(* IEC 61131-3 sources: JingjiangMoonbox/Application/Application/任务列表/CommTask/PRG_COMM, 7 files *)

(* ---- Action_gLink_II_Input.st ---- *)
(*@CES
Name=Action_gLink_II_Input
Type=Action
TypeGuid=8ac092e5-3128-4e26-9e7e-11016c6684f2
Guid=1dfcb6d0-4c04-4e1c-b741-2802373335cf
HasDeclaration=False
HasImplementation=True
*)
{DECLARATION}

{IMPLEMENTATION}
FOR iN:=1 TO MAX_UNIT_NUM BY 1 DO
	pstStUnitParam_Save:= ADR(g_stStSysParam.astStUnitParam_Save[iN]);
	pstStUnitParam_UnSave:= ADR(g_stStSysParam.astStUnitParam_UnSave[iN]);
	//xi.hy2026.5.9.114008
	pstStRSVUnitParam_UnSave:=ADR(g_stStSysParam.astStRSV_UnitParam_UnSave[iN]);

	astStParam_Mailbox_snd[iN].dwSemaphore:= SEMA_DOWNLOAD;
	astStParam_Mailbox_snd[iN].iGateSa:= pstStUnitParam_Save^.iGateSa;
	astStParam_Mailbox_snd[iN].iGateSaEx:= pstStUnitParam_Save^.iGateSaEx;
	astStParam_Mailbox_snd[iN].rAdjust_V:= pstStUnitParam_Save^.rAdj_V;
	astStParam_Mailbox_snd[iN].rAdjust_H:= pstStUnitParam_Save^.rAdj_H;
	astStParam_Mailbox_snd[iN].dwFlag_Ctl:= pstStUnitParam_Save^.dwFlag_Ctl;
	astStParam_Mailbox_snd[iN].dwFlag_Sts:= pstStUnitParam_Save^.dwFlag_Sts;
	//2026.04.08.193624//wButtonFun_Lamp赋值
	pstStUnitParam_Save^.wButtonFun_Lamp.0:=g_astStIOMap_Axis_FE[iN].o_xLamp_Linkage;
	pstStUnitParam_Save^.wButtonFun_Lamp.3:=g_astStIOMap_Axis_FE[iN].o_xLamp_Inch;
	pstStUnitParam_Save^.wButtonFun_Lamp.4:=g_astStIOMap_Axis_FE[iN].o_xLamp_Press;
	pstStUnitParam_Save^.wButtonFun_Lamp.2:=FALSE;
	pstStUnitParam_Save^.wButtonFun_Lamp.5:=FALSE;
	pstStUnitParam_Save^.wButtonFun_Lamp.6:=FALSE;
	//pstStUnitParam_Save^.wButtonFun_Lamp.7:=FALSE;
	pstStUnitParam_Save^.wButtonFun_Lamp.8:=g_astStIOMap_Axis_Extra_FE[iN].o_xRel_TurnoverFilmAgency;
	pstStUnitParam_Save^.wButtonFun_Lamp.9:=FALSE;
	pstStUnitParam_Save^.wButtonFun_Lamp.10:=FALSE;
	pstStUnitParam_Save^.wButtonFun_Lamp.11:=FALSE;
	pstStUnitParam_Save^.wButtonFun_Lamp.12:=FALSE;
	pstStUnitParam_Save^.wButtonFun_Lamp.13:=g_stStSysParam.astStGrpParam_UnSave[1].xFlag_Print OR g_stStSysParam.astStGrpParam_UnSave[1].xFlag_Ink;
	pstStUnitParam_Save^.wButtonFun_Lamp.14:=g_stStSysParam.astStGrpParam_UnSave[1].xFlag_Stop OR g_stStSysParam.astStGrpParam_UnSave[1].xFlag_Stoping;
	astStParam_Mailbox_snd[iN].wButtonFun_Lamp:= pstStUnitParam_Save^.wButtonFun_Lamp;

//	astStParam_Mailbox_snd[iN].wButtonFun_Lamp:= pstStUnitParam_Save^.wButtonFun_Lamp;
	astStParam_Mailbox_snd[iN].wSwitchFun:= pstStUnitParam_Save^.wSwitchFun;
	astStParam_Mailbox_snd[iN].rStep_Pressure_Prn_Net:= pstStUnitParam_Save^.rStep_Pressure_Prn_Net;
	astStParam_Mailbox_snd[iN].rLong_Step_Roller_Pressure:= pstStUnitParam_Save^.rLong_Step_Roller_Pressure;
	astStParam_Mailbox_snd[iN].rShort_Step_Roller_Pressure:= pstStUnitParam_Save^.rShort_Step_Roller_Pressure;
	astStParam_Mailbox_snd[iN].wAirInletWindDoorValue:= pstStUnitParam_Save^.byHotBlower_AO;
	astStParam_Mailbox_snd[iN].wAirExhaustWindDoorValue:= pstStUnitParam_Save^.wAirExhaustWindDoorValue;
	astStParam_Mailbox_snd[iN].wAirReturnWindDoorValue:= pstStUnitParam_Save^.wAirReturnWindDoorValue;
	adwCtlBits_UnitBaseCraft_Temp[iN].0 := pstStUnitParam_Save^.xSwitch_ScraperAuto			;//: BIT;(*刮刀手自动-bit0*)
	adwCtlBits_UnitBaseCraft_Temp[iN].1 := pstStUnitParam_Save^.xSwitch_ScraperOn			;//: BIT;(*刮刀开关bit1*)
	adwCtlBits_UnitBaseCraft_Temp[iN].2 := pstStUnitParam_Save^.xInterver_ScraperRun		;//: BIT;(*刮刀开关bit2*)
	adwCtlBits_UnitBaseCraft_Temp[iN].3 := pstStUnitParam_Save^.xRsv_BIT3					;//: BIT;(*BIT3预留*)
	adwCtlBits_UnitBaseCraft_Temp[iN].4 := pstStUnitParam_Save^.xSwitch_InkRollerAuto		;//: BIT;(*递墨辊手自动bit4*)
	adwCtlBits_UnitBaseCraft_Temp[iN].5 := pstStUnitParam_Save^.xSwitch_InkRollerCW			;//: BIT;(*递墨辊正转bit5*)
	adwCtlBits_UnitBaseCraft_Temp[iN].6 := pstStUnitParam_Save^.xSwitch_InkRollerCCW		;//: BIT;(*递墨辊反转bit6*)
	adwCtlBits_UnitBaseCraft_Temp[iN].7 := pstStUnitParam_Save^.xInterver_InkRollerRun		;//: BIT;(*递墨辊运行bit7*)
	adwCtlBits_UnitBaseCraft_Temp[iN].8 := pstStUnitParam_Save^.xSwitch_HotWindOn			;//: BIT;(*热风开关bit8*)
	adwCtlBits_UnitBaseCraft_Temp[iN].9 := pstStUnitParam_Save^.xInterver_HotWindRun		;//: BIT;(*热风1运行bit9*)
	adwCtlBits_UnitBaseCraft_Temp[iN].10:= pstStUnitParam_Save^.xRsv_BIT10					;//: BIT;(*BIT10预留*)
	adwCtlBits_UnitBaseCraft_Temp[iN].11:= pstStUnitParam_Save^.xRsv_BIT11					;//: BIT;(*BIT11预留*)
	adwCtlBits_UnitBaseCraft_Temp[iN].12:= pstStUnitParam_Save^.xSwitch_HotWindOn_II		;//: BIT;(*热风开关bit12*)
	adwCtlBits_UnitBaseCraft_Temp[iN].13:= pstStUnitParam_Save^.xInterver_HotWindRun_II		;//: BIT;(*热风1运行bit13*)
	adwCtlBits_UnitBaseCraft_Temp[iN].14:= pstStUnitParam_Save^.xRsv_BIT14					;//: BIT;(*BIT14预留*)
	adwCtlBits_UnitBaseCraft_Temp[iN].15:= pstStUnitParam_Save^.xRsv_BIT15					;//: BIT;(*BIT15预留*)
	adwCtlBits_UnitBaseCraft_Temp[iN].16:= pstStUnitParam_Save^.xSwitch_HeatingMode_Water	;//: BIT;(*水加热开关bit16*)
	adwCtlBits_UnitBaseCraft_Temp[iN].17:= pstStUnitParam_Save^.xSwitch_HeatingMode_Ele		;//: BIT;(*电加热开关bit17*)
	adwCtlBits_UnitBaseCraft_Temp[iN].18:= pstStUnitParam_Save^.xSwitch_Heating_I			;//: BIT;(*加热I档bit18*)
	adwCtlBits_UnitBaseCraft_Temp[iN].19:= pstStUnitParam_Save^.xSwitch_Heating_II			;//: BIT;(*加热II档bit19*)
	adwCtlBits_UnitBaseCraft_Temp[iN].20:= pstStUnitParam_Save^.xSwitch_Heating_III			;//: BIT;(*加热III档bit20*)
	adwCtlBits_UnitBaseCraft_Temp[iN].21:= pstStUnitParam_Save^.xRsv_BIT21					;//: BIT;(*BIT21预留*)
	adwCtlBits_UnitBaseCraft_Temp[iN].22:= pstStUnitParam_Save^.xRsv_BIT22					;//: BIT;(*BIT22预留*)
	adwCtlBits_UnitBaseCraft_Temp[iN].23:= pstStUnitParam_Save^.xErrReset_Scraper			;//: BIT;(*刮刀故障复位bit23*)
	adwCtlBits_UnitBaseCraft_Temp[iN].24:= pstStUnitParam_Save^.xErrReset_InkRoller			;//: BIT;(*递墨故障复位bit24*)
	adwCtlBits_UnitBaseCraft_Temp[iN].25:= pstStUnitParam_Save^.xErrReset_Hotwind			;//: BIT;(*热风故障复位bit25*)
	adwCtlBits_UnitBaseCraft_Temp[iN].26:= pstStUnitParam_Save^.xErrReset_Hotwind_II		;//: BIT;(*热风2故障复位bit26*)
	adwCtlBits_UnitBaseCraft_Temp[iN].27:= pstStUnitParam_Save^.xErrReset_ExhAir			;//: BIT;(*排风故障复位bit27*)
	adwCtlBits_UnitBaseCraft_Temp[iN].28:= pstStUnitParam_Save^.xSwitch_ExhAir				;//: BIT;(*排风开关bit28*)
	adwCtlBits_UnitBaseCraft_Temp[iN].29:= pstStUnitParam_Save^.xInterver_ExhAir			;//: BIT;(*排风运行bit29*)
	adwCtlBits_UnitBaseCraft_Temp[iN].30:= pstStUnitParam_Save^.xRsv_BIT30					;//: BIT;(*BIT30预留*)
	adwCtlBits_UnitBaseCraft_Temp[iN].31:= pstStUnitParam_Save^.xSwitch_Coolwind			;//: BIT;(*冷风开关*)

	astStParam_Mailbox_snd[iN].dwCtlBits_UnitBaseCraft:= adwCtlBits_UnitBaseCraft_Temp[iN];
	astStParam_Mailbox_snd[iN].wHz_UnitInkRoller_ManuallySet:= REAL_TO_WORD(pstStUnitParam_Save^.rHz_UnitInkRoller_ManuallySet*100.0);
	astStParam_Mailbox_snd[iN].wCoeff_UnitInkRoller_Auto:= REAL_TO_WORD(pstStUnitParam_Save^.rCoeff_UnitInkRoller_Auto*100.0);
	astStParam_Mailbox_snd[iN].wHz_UnitScraper_ManuallySet:= REAL_TO_WORD(pstStUnitParam_Save^.rHz_UnitScraper_ManuallySet*100.0)		  ;
	astStParam_Mailbox_snd[iN].wCoeff_UnitScraper_Auto:= REAL_TO_WORD(pstStUnitParam_Save^.rCoeff_UnitScraper_Auto*100.0)			     ;
	astStParam_Mailbox_snd[iN].wHz_UnitHotWind:= REAL_TO_WORD(pstStUnitParam_Save^.rHz_UnitHotWind_ManuallySet*100.0)		  ;
	astStParam_Mailbox_snd[iN].wHz_UnitHotWind_2:= REAL_TO_WORD(pstStUnitParam_Save^.rHz_UnitHotWind_2_ManuallySet*100.0)		;
	astStParam_Mailbox_snd[iN].wSV_UnitTemCtl:= REAL_TO_WORD(pstStUnitParam_Save^.rSV_UnitTemCtl*100.0)						           ;
	astStParam_Mailbox_snd[iN].wUnit_output_I:= pstStUnitParam_UnSave^.wUnit_output_I;
	astStParam_Mailbox_snd[iN].wUnit_output_II:= pstStUnitParam_UnSave^.wUnit_output_II;
	astStParam_Mailbox_snd[iN].bySignalSelect:= pstStUnitParam_Save^.bySignalSelect;
	astStParam_Mailbox_snd[iN].rOffset_T1:= pstStUnitParam_Save^.rOffset_T1;
	astStParam_Mailbox_snd[iN].rSource_Light_T1:= pstStUnitParam_Save^.rSource_Light_T1;
	astStParam_Mailbox_snd[iN].rBias_T1:= pstStUnitParam_Save^.rBias_T1;
	astStParam_Mailbox_snd[iN].rBrightness_Light_T1:= pstStUnitParam_Save^.rBrightness_Light_T1;
	astStParam_Mailbox_snd[iN].rOffset_T2:= pstStUnitParam_Save^.rOffset_T2;
	astStParam_Mailbox_snd[iN].rSource_Light_T2:= pstStUnitParam_Save^.rSource_Light_T2;
	astStParam_Mailbox_snd[iN].rBias_T2:= pstStUnitParam_Save^.rBias_T2;
	astStParam_Mailbox_snd[iN].rBrightness_Light_T2:= pstStUnitParam_Save^.rBrightness_Light_T2;

	astStParam_Mailbox_snd[iN].wSlaveBtn_HMI.0:= pstStUnitParam_UnSave^.adwPressureMotor_Move[1].0;//版辊操作侧靠近
	astStParam_Mailbox_snd[iN].wSlaveBtn_HMI.1:= pstStUnitParam_UnSave^.adwPressureMotor_Move[1].1;//版辊操作侧远离
	astStParam_Mailbox_snd[iN].wSlaveBtn_HMI.2:= pstStUnitParam_UnSave^.adwPressureMotor_Move[1].4;//版辊平行靠近
	astStParam_Mailbox_snd[iN].wSlaveBtn_HMI.3:= pstStUnitParam_UnSave^.adwPressureMotor_Move[1].5; //版辊平行远离
	astStParam_Mailbox_snd[iN].wSlaveBtn_HMI.4:= pstStUnitParam_UnSave^.adwPressureMotor_Move[1].2;//版辊传动侧靠近
	astStParam_Mailbox_snd[iN].wSlaveBtn_HMI.5:= pstStUnitParam_UnSave^.adwPressureMotor_Move[1].3;//版辊传动侧远离

	//2026.02.10.143913|新增
	astStParam_Mailbox_snd[iN].wSlaveBtn_HMI.15:= pstStUnitParam_UnSave^.adwPressureMotor_Move[1].10; //版辊合压
	astStParam_Mailbox_snd[iN].wSlaveBtn_HMI2.0:= pstStUnitParam_UnSave^.adwPressureMotor_Move[1].8;//版辊离压
	astStParam_Mailbox_snd[iN].wSlaveBtn_HMI2.3:= pstStUnitParam_UnSave^.adwPressureMotor_Move[1].9;//版辊换版
	//2026.02.23.151133 新增 Hou.N
	astStParam_Mailbox_snd[iN].wSlaveBtn_HMI2.5:= pstStUnitParam_UnSave^.adwPressureMotor_Move[1].14;//自动换版
	astStParam_Mailbox_snd[iN].wSlaveBtn_HMI2.6:= pstStUnitParam_UnSave^.adwPressureMotor_Move[1].15;//版辊换版
	astStParam_Mailbox_snd[iN].wSlaveBtn_HMI2.7:= pstStUnitParam_UnSave^.adwPressureMotor_Move[1].19;//显示换版状态

	astStParam_Mailbox_snd[iN].wSlaveBtn_HMI.6:= pstStUnitParam_UnSave^.adwPressureMotor_Move[2].0;//网辊操作侧靠近
	astStParam_Mailbox_snd[iN].wSlaveBtn_HMI.7:= pstStUnitParam_UnSave^.adwPressureMotor_Move[2].1;//网辊操作侧远离
	astStParam_Mailbox_snd[iN].wSlaveBtn_HMI.8:= pstStUnitParam_UnSave^.adwPressureMotor_Move[2].4;//网辊平行靠近
	astStParam_Mailbox_snd[iN].wSlaveBtn_HMI.9:= pstStUnitParam_UnSave^.adwPressureMotor_Move[2].5;//网辊平行远离
	astStParam_Mailbox_snd[iN].wSlaveBtn_HMI.10:= pstStUnitParam_UnSave^.adwPressureMotor_Move[2].2;//网辊传动侧靠近
	astStParam_Mailbox_snd[iN].wSlaveBtn_HMI.11:= pstStUnitParam_UnSave^.adwPressureMotor_Move[2].3;//网辊传动侧远离

	astStParam_Mailbox_snd[iN].wSlaveBtn_HMI2.1:= pstStUnitParam_UnSave^.adwPressureMotor_Move[2].10;//网辊合压
	astStParam_Mailbox_snd[iN].wSlaveBtn_HMI2.2:= pstStUnitParam_UnSave^.adwPressureMotor_Move[2].8;//网辊离压
	astStParam_Mailbox_snd[iN].wSlaveBtn_HMI2.4:= pstStUnitParam_UnSave^.adwPressureMotor_Move[2].9;//网辊换版

	astStParam_Mailbox_snd[iN].wSlaveBtn_HMI.12:=pstStUnitParam_UnSave^.adwPressureMotor_Move[1].16;//版辊标定
	astStParam_Mailbox_snd[iN].wSlaveBtn_HMI.13:=pstStUnitParam_UnSave^.adwPressureMotor_Move[2].16;//网辊标定
//2026.03.14.93922
	astStParam_Mailbox_snd[iN].wButtonAndSwitch_ChaoXu.1:=pstStUnitParam_Save^.wButtonAndSwitch_ChaoXu.1;//网辊锁轴
	astStParam_Mailbox_snd[iN].wButtonAndSwitch_ChaoXu.2:=pstStUnitParam_Save^.wButtonAndSwitch_ChaoXu.2;//充气
	astStParam_Mailbox_snd[iN].wButtonAndSwitch_ChaoXu.3:=pstStUnitParam_Save^.wButtonAndSwitch_ChaoXu.3;//墨盘电磁阀升
	astStParam_Mailbox_snd[iN].wButtonAndSwitch_ChaoXu.4:=pstStUnitParam_Save^.wButtonAndSwitch_ChaoXu.4;//照明
	astStParam_Mailbox_snd[iN].wButtonAndSwitch_ChaoXu.11:=pstStUnitParam_Save^.wButtonAndSwitch_ChaoXu.11;//合压
	astStParam_Mailbox_snd[iN].wButtonAndSwitch_ChaoXu.12:=pstStUnitParam_Save^.wButtonAndSwitch_ChaoXu.12;//离压
	//2026.03.18.112045 新＋
//	astStParam_Mailbox_snd[iN].wButtonAndSwitch_ChaoXu.5:=pstStUnitParam_Save^.wButtonAndSwitch_ChaoXu.5;//显示是否修改版周
//	astStParam_Mailbox_snd[iN].wButtonAndSwitch_ChaoXu.6:=pstStUnitParam_Save^.wButtonAndSwitch_ChaoXu.6;//确认修改版周
	//2025.11.14.172840  | +
// 	IF pstStUnitParam_Save^.wButtonFun_Lamp.0 THEN
// 		g_astStMcgsBtn_HMI[iN].xBtn_Inch:= TRUE;
// 		pstStUnitParam_Save^.wButtonFun_Lamp.0 := FALSE;
// 	END_IF
	astStParam_Mailbox_snd[iN].wState_FiberMove:=pstStRSVUnitParam_UnSave^.wState_FiberMove;

	g_astStMcgsBtn_HMI[iN].xSwitch_Linkage:= pstStUnitParam_Save^.wSwitchFun.0;
	g_astStMcgsBtn_HMI[iN].xSwitch_PressRollAuto:= pstStUnitParam_Save^.wSwitchFun.1;
	//2026.06.03.132225
	g_astStMcgsBtn_HMI[iN].xSwitch_TurnoverFilm:=pstStUnitParam_Save^.wButtonFun_Lamp.7;

//	g_stStSysParam.astStUnitParam_Save[iN].wButtonFun_Lamp.15:= g_astStIOMap_Axis_FE[iN].o_xLamp_Inch;

		astStParam_Mailbox_snd[iN].iStep_Horz_Use:= REAL_TO_INT(g_stStSysParam.astStRSV_UnitParam_UnSave[iN].rStep_Horz*100.0);
		astStParam_Mailbox_snd[iN].wButtonAndSwitch_ChaoXu.14:= g_stStSysParam.astStRSV_UnitParam_UnSave[iN].xBtn_FromHMI_HorMove_M;
		astStParam_Mailbox_snd[iN].wButtonAndSwitch_ChaoXu.13:= g_stStSysParam.astStRSV_UnitParam_UnSave[iN].xBtn_FromHMI_HorMove_G;

		//2026.03.11.101506  Hou.N +
		astStParam_Mailbox_snd[iN].wButtonAndSwitch_ChaoXu.0:=g_stStSysParam.astStRSV_UnitParam_UnSave[iN].xSwitch_Inching_Net;//匀墨
		astStParam_Mailbox_snd[iN].wButtonAndSwitch_ChaoXu.9:=g_stStSysParam.astStRSV_UnitParam_UnSave[iN].xSwitch_Inching_Prn;//版辊单动
		astStParam_Mailbox_snd[iN].wButtonAndSwitch_ChaoXu.10:=g_stStSysParam.astStRSV_UnitParam_UnSave[iN].xSwitch_Inching_Bottom;//底辊单动

		//xi.hy
		astStParam_Mailbox_snd[iN].wState_FiberMove:=pstStRSVUnitParam_UnSave^.wState_FiberMove;
		astStParam_Mailbox_snd[iN].wAlarm_FiberMove:=pstStRSVUnitParam_UnSave^.uiFiberMoveAlarm;
		astStParam_Mailbox_snd[iN].iFiberMoveDistanceIn:=REAL_TO_WORD(pstStRSVUnitParam_UnSave^.rFiberMoveDistanceIn*10);
		astStParam_Mailbox_snd[iN].iPosCur_FiberMove:=	REAL_TO_INT(pstStRSVUnitParam_UnSave^.rFiberMovePosCur*10.0);
		astStParam_Mailbox_snd[iN].iWidth_FindMarkCenter:= REAL_TO_INT(	pstStRSVUnitParam_UnSave^.rWidth_FindMarkCenter*100.0);

		//2026.04.28.133304 xi.hy新增@七号开始
		astStParam_Mailbox_snd[iN].iStsSlave_FiberMove:=pstStRSVUnitParam_UnSave^.iStsSlave_FiberMove;
		//2026.05.28.181703
		astStParam_Mailbox_snd[iN].iFiberMoveBasePosFromSlave:=REAL_TO_INT(pstStRSVUnitParam_UnSave^.rFiberMoveBasePosFromSlave*10.0);

(*2026.5.9.114326
		astStParam_Mailbox_snd[iN].wAccButton_Count		:=g_awAccButton_Count[iN]		;//		: WORD;
		astStParam_Mailbox_snd[iN].wDecButton_Count		:=g_awDecButton_Count[iN]		;//	: WORD;
		astStParam_Mailbox_snd[iN].wUpAdjButton_Count	:=g_awUpAdjButton_Count[iN]	;	//	: WORD;
		astStParam_Mailbox_snd[iN].wDnAdjButton_Count	:=g_awDnAdjButton_Count[iN]	;	//	: WORD;
		astStParam_Mailbox_snd[iN].wLeftAdjButton_Count	:=g_awLeftAdjButton_Count[iN]	;	//		: WORD;
		astStParam_Mailbox_snd[iN].wRightAdjButton_Count	:=g_awRightAdjButton_Count[iN];	//		: WORD;
		astStParam_Mailbox_snd[iN].wAlarmButton_Count:= g_awAlarmButton_Count[iN]		;//	: WORD;
	*)
END_FOR

(* ---- Action_gLink_II_Output.st ---- *)
(*@CES
Name=Action_gLink_II_Output
Type=Action
TypeGuid=8ac092e5-3128-4e26-9e7e-11016c6684f2
Guid=075e8bd3-4afc-466b-b5b0-16bdc62b582f
HasDeclaration=False
HasImplementation=True
*)
{DECLARATION}

{IMPLEMENTATION}
FOR iN:=1 TO MAX_UNIT_NUM BY 1 DO
	pstStUnitParam_Save:= ADR(g_stStSysParam.astStUnitParam_Save[iN]);
	pstStUnitParam_UnSave:= ADR(g_stStSysParam.astStUnitParam_UnSave[iN]);
	//xi.hy2026.5.9.114419
	pstStRSVUnitParam_UnSave:=ADR(g_stStSysParam.astStRSV_UnitParam_UnSave[iN]);
	IF axNeedUpdateParam_Malilbox[iN] THEN
		axNeedUpdateParam_Malilbox[iN]:= FALSE;
		pstStUnitParam_Save^.iGateSa:= astStParam_Mailbox_out[iN].iGateSa                      	;//第一波门位置
		pstStUnitParam_Save^.iGateSaEx:= astStParam_Mailbox_out[iN].iGateSaEx                        ;//第二波门位置
		pstStUnitParam_Save^.rAdj_V:= astStParam_Mailbox_out[iN].rAdjust_V                        ;//纵向版修正量
		pstStUnitParam_Save^.rAdj_H:= astStParam_Mailbox_out[iN].rAdjust_H                        ;//横向版修正量
		pstStUnitParam_Save^.dwFlag_Ctl:= astStParam_Mailbox_out[iN].dwFlag_Ctl                       ;//套色控制标志
		pstStUnitParam_Save^.dwFlag_Sts:= astStParam_Mailbox_out[iN].dwFlag_Sts                       ;//套色状态标志
		pstStUnitParam_Save^.wButtonFun_Lamp:= astStParam_Mailbox_out[iN].wButtonFun_Lamp                  ;//HMI界面按钮及指示灯
		//2026.04.08.195419||2026.5.9.114523
		g_astStMcgsBtn_HMI[iN].xBtn_Inch:=pstStUnitParam_Save^.wButtonFun_Lamp.2;
		g_astStMcgsBtn_HMI[iN].xBtn_Press:=pstStUnitParam_Save^.wButtonFun_Lamp.5;
		g_astStMcgsBtn_HMI[iN].xBtn_UnPress:=pstStUnitParam_Save^.wButtonFun_Lamp.6;
		//g_astStMcgsBtn_HMI[iN].xBtn_TurnoverFilm:=pstStUnitParam_Save^.wButtonFun_Lamp.7;
		g_astStMcgsBtn_HMI[iN].xBtn_Stop:=pstStUnitParam_Save^.wButtonFun_Lamp.9;
		g_astStMcgsBtn_HMI[iN].xBtn_Ink:=pstStUnitParam_Save^.wButtonFun_Lamp.10;
		g_astStMcgsBtn_HMI[iN].xBtn_Print:=pstStUnitParam_Save^.wButtonFun_Lamp.11;
		g_astStMcgsBtn_HMI[iN].xBtn_PreStart:=pstStUnitParam_Save^.wButtonFun_Lamp.12;

		pstStUnitParam_Save^.wSwitchFun:= astStParam_Mailbox_out[iN].wSwitchFun                   ;//界面按钮
		pstStUnitParam_Save^.rStep_Pressure_Prn_Net:= astStParam_Mailbox_out[iN].rStep_Pressure_Prn_Net           ;//版辊网辊按钮步进量
		pstStUnitParam_Save^.rLong_Step_Roller_Pressure:= astStParam_Mailbox_out[iN].rLong_Step_Roller_Pressure       ;//色组压力控制长步进值
		pstStUnitParam_Save^.rShort_Step_Roller_Pressure:= astStParam_Mailbox_out[iN].rShort_Step_Roller_Pressure      ;//色组压力控制短步进值
		pstStUnitParam_Save^.byHotBlower_AO:= WORD_TO_BYTE(astStParam_Mailbox_out[iN].wAirInletWindDoorValue)           ;//进风口风门开度值
		pstStUnitParam_Save^.wAirExhaustWindDoorValue:= astStParam_Mailbox_out[iN].wAirExhaustWindDoorValue         ;//排风口风门开度值
		pstStUnitParam_Save^.wAirReturnWindDoorValue:= astStParam_Mailbox_out[iN].wAirReturnWindDoorValue          ;//回风口风门开度值

		adwCtlBits_UnitBaseCraft_Temp[iN]:= astStParam_Mailbox_out[iN].dwCtlBits_UnitBaseCraft          ;//界面工艺开关及状态

		pstStUnitParam_Save^.xSwitch_ScraperAuto			:= adwCtlBits_UnitBaseCraft_Temp[iN].0 ;//: BIT;(*刮刀手自动-bit0*)
		pstStUnitParam_Save^.xSwitch_ScraperOn			:= adwCtlBits_UnitBaseCraft_Temp[iN].1 ;//: BIT;(*刮刀开关bit1*)
		pstStUnitParam_Save^.xInterver_ScraperRun		:= adwCtlBits_UnitBaseCraft_Temp[iN].2 ;//: BIT;(*刮刀开关bit2*)
		pstStUnitParam_Save^.xRsv_BIT3					:= adwCtlBits_UnitBaseCraft_Temp[iN].3 ;//: BIT;(*BIT3预留*)
		pstStUnitParam_Save^.xSwitch_InkRollerAuto		:= adwCtlBits_UnitBaseCraft_Temp[iN].4 ;//: BIT;(*递墨辊手自动bit4*)
		pstStUnitParam_Save^.xSwitch_InkRollerCW			:= adwCtlBits_UnitBaseCraft_Temp[iN].5 ;//: BIT;(*递墨辊正转bit5*)
		pstStUnitParam_Save^.xSwitch_InkRollerCCW		:= adwCtlBits_UnitBaseCraft_Temp[iN].6 ;//: BIT;(*递墨辊反转bit6*)
		pstStUnitParam_Save^.xInterver_InkRollerRun		:= adwCtlBits_UnitBaseCraft_Temp[iN].7 ;//: BIT;(*递墨辊运行bit7*)
		pstStUnitParam_Save^.xSwitch_HotWindOn			:= adwCtlBits_UnitBaseCraft_Temp[iN].8 ;//: BIT;(*热风开关bit8*)
		pstStUnitParam_Save^.xInterver_HotWindRun		:= adwCtlBits_UnitBaseCraft_Temp[iN].9 ;//: BIT;(*热风1运行bit9*)
		pstStUnitParam_Save^.xRsv_BIT10					:= adwCtlBits_UnitBaseCraft_Temp[iN].10;//: BIT;(*BIT10预留*)
		pstStUnitParam_Save^.xRsv_BIT11					:= adwCtlBits_UnitBaseCraft_Temp[iN].11;//: BIT;(*BIT11预留*)
		pstStUnitParam_Save^.xSwitch_HotWindOn_II		:= adwCtlBits_UnitBaseCraft_Temp[iN].12;//: BIT;(*热风开关bit12*)
		pstStUnitParam_Save^.xInterver_HotWindRun_II		:= adwCtlBits_UnitBaseCraft_Temp[iN].13;//: BIT;(*热风1运行bit13*)
		pstStUnitParam_Save^.xRsv_BIT14					:= adwCtlBits_UnitBaseCraft_Temp[iN].14;//: BIT;(*BIT14预留*)
		pstStUnitParam_Save^.xRsv_BIT15					:= adwCtlBits_UnitBaseCraft_Temp[iN].15;//: BIT;(*BIT15预留*)
		pstStUnitParam_Save^.xSwitch_HeatingMode_Water	:= adwCtlBits_UnitBaseCraft_Temp[iN].16;//: BIT;(*水加热开关bit16*)
		pstStUnitParam_Save^.xSwitch_HeatingMode_Ele		:= adwCtlBits_UnitBaseCraft_Temp[iN].17;//: BIT;(*电加热开关bit17*)
		pstStUnitParam_Save^.xSwitch_Heating_I			:= adwCtlBits_UnitBaseCraft_Temp[iN].18;//: BIT;(*加热I档bit18*)
		pstStUnitParam_Save^.xSwitch_Heating_II			:= adwCtlBits_UnitBaseCraft_Temp[iN].19;//: BIT;(*加热II档bit19*)
		pstStUnitParam_Save^.xSwitch_Heating_III			:= adwCtlBits_UnitBaseCraft_Temp[iN].20;//: BIT;(*加热III档bit20*)
		pstStUnitParam_Save^.xRsv_BIT21					:= adwCtlBits_UnitBaseCraft_Temp[iN].21;//: BIT;(*BIT21预留*)
		pstStUnitParam_Save^.xRsv_BIT22					:= adwCtlBits_UnitBaseCraft_Temp[iN].22;//: BIT;(*BIT22预留*)
		pstStUnitParam_Save^.xErrReset_Scraper			:= adwCtlBits_UnitBaseCraft_Temp[iN].23;//: BIT;(*刮刀故障复位bit23*)
		pstStUnitParam_Save^.xErrReset_InkRoller			:= adwCtlBits_UnitBaseCraft_Temp[iN].24;//: BIT;(*递墨故障复位bit24*)
		pstStUnitParam_Save^.xErrReset_Hotwind			:= adwCtlBits_UnitBaseCraft_Temp[iN].25;//: BIT;(*热风故障复位bit25*)
		pstStUnitParam_Save^.xErrReset_Hotwind_II		:= adwCtlBits_UnitBaseCraft_Temp[iN].26;//: BIT;(*热风2故障复位bit26*)
		pstStUnitParam_Save^.xErrReset_ExhAir			:= adwCtlBits_UnitBaseCraft_Temp[iN].27;//: BIT;(*排风故障复位bit27*)
		pstStUnitParam_Save^.xSwitch_ExhAir				:= adwCtlBits_UnitBaseCraft_Temp[iN].28;//: BIT;(*排风开关bit28*)
		pstStUnitParam_Save^.xInterver_ExhAir			:= adwCtlBits_UnitBaseCraft_Temp[iN].29;//: BIT;(*排风运行bit29*)
		pstStUnitParam_Save^.xRsv_BIT30					:= adwCtlBits_UnitBaseCraft_Temp[iN].30;//: BIT;(*BIT30预留*)
		pstStUnitParam_Save^.xSwitch_Coolwind			:= adwCtlBits_UnitBaseCraft_Temp[iN].31;//: BIT;(*冷风开关*)

		pstStUnitParam_Save^.rHz_UnitInkRoller_ManuallySet:= WORD_TO_REAL(astStParam_Mailbox_out[iN].wHz_UnitInkRoller_ManuallySet)/100.0    ;//递墨辊手动频率
		pstStUnitParam_Save^.rCoeff_UnitInkRoller_Auto:= WORD_TO_REAL(astStParam_Mailbox_out[iN].wCoeff_UnitInkRoller_Auto)/100.0         ;//递墨辊自动系数
		pstStUnitParam_Save^.rHz_UnitScraper_ManuallySet:= WORD_TO_REAL(astStParam_Mailbox_out[iN].wHz_UnitScraper_ManuallySet)/100.0       ;//刮刀手动频率
		pstStUnitParam_Save^.rCoeff_UnitScraper_Auto:= WORD_TO_REAL(astStParam_Mailbox_out[iN].wCoeff_UnitScraper_Auto)/100.0           ;//刮刀自动系数
		pstStUnitParam_Save^.rHz_UnitHotWind_ManuallySet:= WORD_TO_REAL(astStParam_Mailbox_out[iN].wHz_UnitHotWind)/100.0                   ;//热风频率
		pstStUnitParam_Save^.rHz_UnitHotWind_2_ManuallySet:= WORD_TO_REAL(astStParam_Mailbox_out[iN].wHz_UnitHotWind_2)/100.0                 ;//热风2频率
		pstStUnitParam_Save^.rSV_UnitTemCtl:= WORD_TO_REAL(astStParam_Mailbox_out[iN].wSV_UnitTemCtl)/100.0                   ;//加热设定温度
		pstStUnitParam_UnSave^.wUnit_output_I:= astStParam_Mailbox_out[iN].wUnit_output_I                   ;//IO监控输出1
		pstStUnitParam_UnSave^.wUnit_output_II:= astStParam_Mailbox_out[iN].wUnit_output_II                  ;//IO监控输出2
		//xi.hy//增加
		pstStUnitParam_Save^.bySignalSelect:= astStParam_Mailbox_out[iN].bySignalSelect;
		pstStUnitParam_Save^.rOffset_T1:= astStParam_Mailbox_out[iN].rOffset_T1             				;//T1路光纤电眼偏移控制
		pstStUnitParam_Save^.rSource_Light_T1:= astStParam_Mailbox_out[iN].rSource_Light_T1                ;//T1路光纤电眼光源控制
		pstStUnitParam_Save^.rBias_T1:= astStParam_Mailbox_out[iN].rBias_T1								;//T1路光纤电眼偏置控制
		pstStUnitParam_Save^.rBrightness_Light_T1:= astStParam_Mailbox_out[iN].rBrightness_Light_T1        ;//T1路光纤电眼亮度控制

		pstStUnitParam_Save^.rOffset_T2:= astStParam_Mailbox_out[iN].rOffset_T2             				;//T2路光纤电眼偏移控制
		pstStUnitParam_Save^.rSource_Light_T2:= astStParam_Mailbox_out[iN].rSource_Light_T2                ;//T2路光纤电眼光源控制
		pstStUnitParam_Save^.rBias_T2:= astStParam_Mailbox_out[iN].rBias_T2								;//T2路光纤电眼偏置控制
		pstStUnitParam_Save^.rBrightness_Light_T2:= astStParam_Mailbox_out[iN].rBrightness_Light_T2        ;//T2路光纤电眼亮度控制
		//2026.02.05.161226 新增 Hou.N
		pstStUnitParam_UnSave^.adwPressureMotor_Move[1].0:=astStParam_Mailbox_out[iN].wSlaveBtn_HMI.0;//版辊操作侧靠近
		pstStUnitParam_UnSave^.adwPressureMotor_Move[1].1:=astStParam_Mailbox_out[iN].wSlaveBtn_HMI.1;//版辊操作侧远离
		pstStUnitParam_UnSave^.adwPressureMotor_Move[1].4:=astStParam_Mailbox_out[iN].wSlaveBtn_HMI.2;//版辊平行靠近
		pstStUnitParam_UnSave^.adwPressureMotor_Move[1].5:=astStParam_Mailbox_out[iN].wSlaveBtn_HMI.3; //版辊平行远离
		pstStUnitParam_UnSave^.adwPressureMotor_Move[1].2:=astStParam_Mailbox_out[iN].wSlaveBtn_HMI.4;//版辊传动侧靠近
		pstStUnitParam_UnSave^.adwPressureMotor_Move[1].3:=astStParam_Mailbox_out[iN].wSlaveBtn_HMI.5;//版辊传动侧远离

//2026.02.10.143913|新增
		pstStUnitParam_UnSave^.adwPressureMotor_Move[1].16:=astStParam_Mailbox_out[iN].wSlaveBtn_HMI.12; //版辊标定
		pstStUnitParam_UnSave^.adwPressureMotor_Move[2].16:=astStParam_Mailbox_out[iN].wSlaveBtn_HMI.13;//网辊标定
	//	pstStUnitParam_UnSave^.adwPressureMotor_Move[3].16:=astStParam_Mailbox_out[iN].dwSlaveBtn_HMI.14;//张带棍标定

		pstStUnitParam_UnSave^.adwPressureMotor_Move[1].10:=astStParam_Mailbox_out[iN].wSlaveBtn_HMI.15; //版辊合压
		pstStUnitParam_UnSave^.adwPressureMotor_Move[1].8:=astStParam_Mailbox_out[iN].wSlaveBtn_HMI2.0;//版辊离压
		IF  astStParam_Mailbox_out[iN].wSlaveBtn_HMI2.0 OR astStParam_Mailbox_out[iN].wSlaveBtn_HMI.15 THEN
			aiTime1[4]:= aiTime1[4]+1;
		END_IF

		pstStUnitParam_UnSave^.adwPressureMotor_Move[1].9:=astStParam_Mailbox_out[iN].wSlaveBtn_HMI2.3;//版辊换版
	//2026.02.23.133406 新增
		pstStUnitParam_UnSave^.adwPressureMotor_Move[1].14:=astStParam_Mailbox_out[iN].wSlaveBtn_HMI2.5;//自动换版
		pstStUnitParam_UnSave^.adwPressureMotor_Move[1].15:=astStParam_Mailbox_out[iN].wSlaveBtn_HMI2.6;//换版完成
		pstStUnitParam_UnSave^.adwPressureMotor_Move[1].19:=astStParam_Mailbox_out[iN].wSlaveBtn_HMI2.7;//显示换版状态

		pstStUnitParam_UnSave^.adwPressureMotor_Move[2].0:=astStParam_Mailbox_out[iN].wSlaveBtn_HMI.6;//网辊操作侧靠近
		pstStUnitParam_UnSave^.adwPressureMotor_Move[2].1:=astStParam_Mailbox_out[iN].wSlaveBtn_HMI.7;//网辊操作侧远离
		pstStUnitParam_UnSave^.adwPressureMotor_Move[2].4:=astStParam_Mailbox_out[iN].wSlaveBtn_HMI.8;//网辊平行靠近
		pstStUnitParam_UnSave^.adwPressureMotor_Move[2].5:=astStParam_Mailbox_out[iN].wSlaveBtn_HMI.9;//网辊平行远离
		pstStUnitParam_UnSave^.adwPressureMotor_Move[2].2:=astStParam_Mailbox_out[iN].wSlaveBtn_HMI.10;//网辊传动侧靠近
		pstStUnitParam_UnSave^.adwPressureMotor_Move[2].3:=astStParam_Mailbox_out[iN].wSlaveBtn_HMI.11;//网辊传动侧远离

		IF astStParam_Mailbox_out[iN].wSlaveBtn_HMI.6 THEN
			g_aiTestBtn[In]:= g_aiTestBtn[In] +1;
		END_IF
		IF astStParam_Mailbox_out[iN].wSlaveBtn_HMI.7 THEN
			g_aiTestBtn1[In]:= g_aiTestBtn1[In] +1;
		END_IF

		IF astStParam_Mailbox_out[iN].wSlaveBtn_HMI.8 THEN
			g_aiTestBtn2[In]:= g_aiTestBtn2[In] +1;
		END_IF

		IF astStParam_Mailbox_out[iN].wSlaveBtn_HMI.9 THEN
			g_aiTestBtn3[In]:= g_aiTestBtn3[In] +1;
		END_IF

		IF astStParam_Mailbox_out[iN].wSlaveBtn_HMI.10  THEN
			g_aiTestBtn4[In]:= g_aiTestBtn4[In] +1;
		END_IF
		IF astStParam_Mailbox_out[iN].wSlaveBtn_HMI.11 THEN
			g_aiTestBtn5[In]:= g_aiTestBtn5[In] +1;
		END_IF

	//2026.02.10.143913|新增
		pstStUnitParam_UnSave^.adwPressureMotor_Move[2].10:=astStParam_Mailbox_out[iN].wSlaveBtn_HMI2.1;//网辊合压
		pstStUnitParam_UnSave^.adwPressureMotor_Move[2].8:=astStParam_Mailbox_out[iN].wSlaveBtn_HMI2.2;//网辊离压
		pstStUnitParam_UnSave^.adwPressureMotor_Move[2].9:=astStParam_Mailbox_out[iN].wSlaveBtn_HMI2.4;//网辊换版

	//2026.03.11.101506 Hou.N +
		g_stStSysParam.astStRSV_UnitParam_UnSave[iN].xSwitch_Inching_Net:=astStParam_Mailbox_out[iN].wButtonAndSwitch_ChaoXu.0;//匀墨
		g_stStSysParam.astStRSV_UnitParam_UnSave[iN].xSwitch_Inching_Prn:=astStParam_Mailbox_out[iN].wButtonAndSwitch_ChaoXu.9;//版辊单动
		g_stStSysParam.astStRSV_UnitParam_UnSave[iN].xSwitch_Inching_Bottom:=astStParam_Mailbox_out[iN].wButtonAndSwitch_ChaoXu.10;//底辊单动

		g_stStSysParam.astStRSV_UnitParam_UnSave[iN].rStep_Horz:= INT_TO_REAL(astStParam_Mailbox_out[iN].iStep_Horz_Use)/100.0;
		g_stStSysParam.astStRSV_UnitParam_UnSave[iN].xBtn_FromHMI_HorMove_M:= astStParam_Mailbox_out[iN].wButtonAndSwitch_ChaoXu.14;
		g_stStSysParam.astStRSV_UnitParam_UnSave[iN].xBtn_FromHMI_HorMove_G:= astStParam_Mailbox_out[iN].wButtonAndSwitch_ChaoXu.13;

		pstStUnitParam_Save^.wButtonAndSwitch_ChaoXu.1:=astStParam_Mailbox_out[iN].wButtonAndSwitch_ChaoXu.1;//网辊锁轴
		pstStUnitParam_Save^.wButtonAndSwitch_ChaoXu.2:=astStParam_Mailbox_out[iN].wButtonAndSwitch_ChaoXu.2;//充气
		pstStUnitParam_Save^.wButtonAndSwitch_ChaoXu.3:=astStParam_Mailbox_out[iN].wButtonAndSwitch_ChaoXu.3;//墨盘电磁阀升
		pstStUnitParam_Save^.wButtonAndSwitch_ChaoXu.4:=astStParam_Mailbox_out[iN].wButtonAndSwitch_ChaoXu.4;//照明
		pstStUnitParam_Save^.wButtonAndSwitch_ChaoXu.11:=astStParam_Mailbox_out[iN].wButtonAndSwitch_ChaoXu.11;//合压
		pstStUnitParam_Save^.wButtonAndSwitch_ChaoXu.12:=astStParam_Mailbox_out[iN].wButtonAndSwitch_ChaoXu.12;//离压

	pstStUnitParam_Save^.wButtonAndSwitch_ChaoXu.5:= FALSE;
	pstStUnitParam_Save^.wButtonAndSwitch_ChaoXu.6:= FALSE;
	pstStUnitParam_Save^.wButtonAndSwitch_ChaoXu.7:= FALSE;

		//xi.hy
		//IF(awState_FiberMove_bak[iN]<>astStParam_Mailbox_out[iN].wState_FiberMove) THEN
			pstStRSVUnitParam_UnSave^.wState_FiberMove:=astStParam_Mailbox_out[iN].wState_FiberMove;
		//	awState_FiberMove_bak[iN]:=astStParam_Mailbox_out[iN].wState_FiberMove;
	//	END_IF

		pstStRSVUnitParam_UnSave^.uiFiberMoveAlarm:=astStParam_Mailbox_out[iN].wAlarm_FiberMove;
		pstStRSVUnitParam_UnSave^.rFiberMoveDistanceIn:=INT_TO_REAL(astStParam_Mailbox_out[iN].iFiberMoveDistanceIn)/10.0;
		pstStRSVUnitParam_UnSave^.rFiberMovePosCur:=INT_TO_REAL(astStParam_Mailbox_out[iN].iPosCur_FiberMove)/10.0;
		pstStRSVUnitParam_UnSave^.rWidth_FindMarkCenter:=INT_TO_REAL(astStParam_Mailbox_out[iN].iWidth_FindMarkCenter)/100.0;

		//2026.04.28.133209 xi.hy新增@七号开始
		pstStRSVUnitParam_UnSave^.iStsSlave_FiberMove:=astStParam_Mailbox_out[iN].iStsSlave_FiberMove;
		//2026.05.28.181905
		pstStRSVUnitParam_UnSave^.rFiberMoveBasePosFromSlave:=INT_TO_REAL(astStParam_Mailbox_out[iN].iFiberMoveBasePosFromSlave)/10.0;

IF  astStParam_Mailbox_out[iN].wButtonAndSwitch_ChaoXu.13 THEN
	aiTime[In]:= aiTime[In] +1;
END_IF
	//2026.02.05.195231
	IF pstStUnitParam_Save^.wButtonAndSwitch_ChaoXu.11 THEN
		g_astStMcgsBtn_HMI[iN].xBtn_Press:= TRUE;
		pstStUnitParam_Save^.wButtonAndSwitch_ChaoXu.11 := FALSE;
	END_IF
	IF pstStUnitParam_Save^.wButtonAndSwitch_ChaoXu.12 THEN
		g_astStMcgsBtn_HMI[iN].xBtn_UnPress:= TRUE;
		pstStUnitParam_Save^.wButtonAndSwitch_ChaoXu.12 := FALSE;
	END_IF

		SysMemSet(adr(astStParam_Mailbox_out[iN]),0,sizeof(astStParam_Mailbox_out[iN]));
	END_IF

	//2025.11.14.172840  | + |延时6个周期请标志
	IF g_astStMcgsBtn_HMI[iN].xBtn_Inch THEN
		aiCntInch[iN] := aiCntInch[iN] + 1;
		IF aiCntInch[iN] > 5 THEN
			aiCntInch[iN] := 0;
			g_astStMcgsBtn_HMI[iN].xBtn_Inch := FALSE;
		END_IF
	ELSE
		aiCntInch[iN] := 0;
	END_IF

	IF g_astStMcgsBtn_HMI[iN].xBtn_Press THEN
		aiCntPress[iN] := aiCntPress[iN] + 1;
		IF aiCntPress[iN] > 10 THEN
			aiCntPress[iN] := 0;
			g_astStMcgsBtn_HMI[iN].xBtn_Press := FALSE;
		END_IF
	ELSE
		aiCntPress[iN] := 0;
	END_IF

	IF g_astStMcgsBtn_HMI[iN].xBtn_UnPress THEN
		aiCntUnPress[iN] := aiCntUnPress[iN] + 1;
		IF aiCntUnPress[iN] > 10 THEN
			aiCntUnPress[iN] := 0;
			g_astStMcgsBtn_HMI[iN].xBtn_UnPress := FALSE;
		END_IF
	ELSE
		aiCntUnPress[iN] := 0;
	END_IF

	//2026.08.06.203030+
	IF g_astStMcgsBtn_HMI[iN].xBtn_Stop THEN
		aiCntStop[iN] := aiCntStop[iN] + 1;
		IF aiCntStop[iN] > 5 THEN
			aiCntStop[iN] := 0;
			g_astStMcgsBtn_HMI[iN].xBtn_Stop := FALSE;
		END_IF
	ELSE
		aiCntStop[iN] := 0;
	END_IF

END_FOR

(* ---- Action_GLINKII_COMM.st ---- *)
(*@CES
Name=Action_GLINKII_COMM
Type=Action
TypeGuid=8ac092e5-3128-4e26-9e7e-11016c6684f2
Guid=d0921674-03aa-48cd-942a-bf6130ef7c95
HasDeclaration=False
HasImplementation=True
*)
{DECLARATION}

{IMPLEMENTATION}
(* ************************************************** *)
(* 命令轮询队列的初始化 *)
(* ************************************************** *)
IF NOT xFlag_CmdQueueInitialized THEN
	FOR iN:=1 TO MAX_UNIT_NUM BY 1 DO
		astStUnitCmdQueue[iN].aiCmdId[1]:= 91;
		astStUnitCmdQueue[iN].aiCmdId[2]:= 92;
		astStUnitCmdQueue[iN].aiCmdId[3]:= 93;
		astStUnitCmdQueue[iN].aiCmdId[4]:= 94;
		astStUnitCmdQueue[iN].aiCmdId[5]:= 95;

		astStUnitCmdQueue[iN].byCmdNum:= 5;

		astStUnitCmdQueue[iN].byCmdIdx:= 1;
	END_FOR
	xFlag_CmdQueueInitialized:= TRUE;
	tmPduSnt_LastTime:= tmCURR;
ELSE
	;
END_IF
(* 有个内存需要申请 *)
IF pastStParam_Mailbox_proof=0 THEN
	pastStParam_Mailbox_proof:= SysMemAllocData('',SIZEOF(pastStParam_Mailbox_proof^),ADR(udiresult));
ELSE
	;
END_IF
(* h/
/pdu通讯/(广播命令)
/每次调用对列表中所有的站只处理各自的1条广播命令
*)

tmCURR:= TIME();
IF (tmCURR-tmPduSnt_LastTime)>=TIMEOUTS_PDU_CMD_CHG THEN(* 时间到/开始处理pdu命令轮询 *)
	FOR iN:=1 TO MAX_UNIT_NUM BY 1 DO(* 为了保证让所有的都能同步轮询命令id/这里把所有色组都循环上 *)
		iUnitId:= iN;(*通讯轴号也需要根据后续系统配置处理*)
		pstStUnitCmdQueue_Tmp:= ADR(astStUnitCmdQueue[iUnitId]);
		iGrpId := KS_GetGrpIdByAxisId(iUnitId,ADR(g_stStSysParam),ADR(iAxisTypeId));
		iStationId := g_stStSysParam.stStSysParam_UnSave.aiStationList_UnitController[iN];
		IF pstStUnitCmdQueue_Tmp<>0 AND
			KS_IsValidStationNR(iStationId) AND
			(iGrpId=1 OR iGrpId=2) AND (* 已经明确分配AB系 *)
			iStationId<>g_stStStationInfo_KS.iSid_Device THEN(*2024.1.3.200526/+ *)

			byIDX_Tmp:= pstStUnitCmdQueue_Tmp^.byCmdIdx;
			byMAX_Tmp:= pstStUnitCmdQueue_Tmp^.byCmdNum;
			IF (byIDX_Tmp>=1 AND byIDX_Tmp<=byMAX_Tmp) AND
				(byMAX_Tmp<=MAX_CMD_NUM_PDU) THEN(* 命令轮询范围有效 *)
				iRtn:=
				KS_FillUnitPduCmd_DN(
					iUnitId,
					iGrpId,
					astStUnitCmdQueue[iUnitId].aiCmdId[byIDX_Tmp],
					wAxis_RollerDn,
					wAxis_Alarm_Prn,
					wComplexFlag_AxisInching,
					wComplexFlag_Linkage,
					ADR(g_stStSysParam),
					ADR(abyBuf_PduCmd_snd));
				IF iRtn=0 THEN
					dwOFST:= 0;
					dwOFST.14:= TRUE;(* 绝对地址访问 *)

					(* pdu发送 *)
					iRtn:=
					GTN_RN_UserPCWrNetFPGA(
						1,(*卡号，先只写1*)
						1,(*总线ID，第一套等环网写1，第二套等环网写2*)
						iStationId,(*物理站号*)
						ADR(abyBuf_PduCmd_snd),	(*有效数据*)
						DWORD_TO_WORD(dwOFST),(*地址*)
						KS_GetNumOfDwordUsed(SIZEOF(abyBuf_PduCmd_snd)) );
					IF iRtn<>0 THEN
						(*写日志2023.3.31.095202*)
						;
					ELSE
						//2026.04.03.114245PDU只要通讯正常，Mailbox不需要考虑强制10s更新参数
						atmUnitMailboxLastSynchronized[iUnitId]:= tmCURR;

					END_IF
				ELSE
					;
				END_IF
				IF byIDX_Tmp>=byMAX_Tmp THEN
					byIDX_Tmp:=1;
				ELSE
					byIDX_Tmp:= byIDX_Tmp+1;
				END_IF
				pstStUnitCmdQueue_Tmp^.byCmdIdx:= byIDX_Tmp;
			ELSE
				pstStUnitCmdQueue_Tmp^.byCmdIdx:= 1;
			END_IF
		ELSE
			;
		END_IF
	END_FOR
	tmPduSnt_LastTime:= tmCURR;(* 更新时间戳 *)
ELSE
	;
END_IF

(* ************************************************** *)
(* 开始处理mailbox通讯 *)
(* MAILbox处理机制: *)
(* 按照16个色组(MAX_UNIT_NUM)来均分8k区域/每区域512字节 *)
(* 按照最大Mailbox单包最大字节480字节进行约束 *)
(* 每个区域都是按照轴进行分配的 *)
(* ************************************************** *)
FOR iN:=1 TO MAX_UNIT_NUM BY 1 DO
	iUnitId:= iN;
	dwOFST:= INT_TO_DWORD((iUnitId-1))*INT_TO_DWORD(MAILBOX_PKG_MAX_BYTES);
	iStationId := g_stStSysParam.stStSysParam_UnSave.aiStationList_UnitController[iUnitId];
	pstStUnitParam_Save:= ADR(g_stStSysParam.astStUnitParam_Save[iUnitId]);
	pstStUnitParam_UnSave:= ADR(g_stStSysParam.astStUnitParam_UnSave[iUnitId]);

	IF pstStUnitParam_Save<>0 AND(* 色组id访问有效 *)
		KS_IsValidStationNR(iStationId) AND(*2024.1.3.200526/+ *)
		iUnitId<=MIN(MAX_UNIT_NUM,g_stStSysParam.stStSysParam_Save.iUnitMaxNum) AND
		iStationId<>g_stStStationInfo_KS.iSid_Device THEN(* 色组有效范围内/循环最少的数量/2023.11.22.102021/han.dp *)
														//增加判断-不与自身站通讯
		(* 本地读取/1次多读1点/万一是需要的就不用再读了 *)
		pDataTest:= adr(abyBuf_MailboxPkg_rcv);
		iRtn:= GTN_RN_DevicePcMailRd(
								1,
								1,
								0,
								ADR(abyBuf_MailboxPkg_rcv),
								DWORD_TO_WORD(dwOFST),
								KS_GetNumOfDwordUsed(SIZEOF(pstStParam_Mailbox_Tmp^)),
								RN_ARD);
		//2023.12.26.163244通讯长度改为实际长度2023.12.26.163251
		(* 套用协议/2021.12.21.114854/hdp *)
		pstStParam_Mailbox_Tmp:= ADR(abyBuf_MailboxPkg_rcv);
		(* gt指令执行成功且协议套用成功/2021.12.21.114917/hdp *)
		IF iRtn=0 AND pstStParam_Mailbox_Tmp<>0 THEN
			CASE pstStParam_Mailbox_Tmp^.dwSemaphore OF
			SEMA_UPLOAD:(* 来自从站的数据更新/没什么问题就同步到本地数据结构中 *)

				(* 判断一下参数的合理性/如果有问题/强行同步到从站去 *)
				IF (pstStParam_Mailbox_Tmp^.iGateSa>=0 AND pstStParam_Mailbox_Tmp^.iGateSa<=3999) AND
					(pstStParam_Mailbox_Tmp^.iGateSaEx>=0 AND pstStParam_Mailbox_Tmp^.iGateSaEx<=3999) AND
					(pstStParam_Mailbox_Tmp^.rAdjust_V>=-80.00 AND pstStParam_Mailbox_Tmp^.rAdjust_V<=80.00) AND
					(pstStParam_Mailbox_Tmp^.rAdjust_H>=-20.00 AND pstStParam_Mailbox_Tmp^.rAdjust_H<=20.00) AND
					(NOT (pstStParam_Mailbox_Tmp^.wSV_UnitTemCtl=0 AND pstStUnitParam_Save^.rSV_UnitTemCtl<>0))
					 THEN//参数
							(*2023.12.26.150253增加保护-设定温度不会主动设定为0取*)
							(* 重要的几个参数检查/合法通过后 *)
					axNeedUpdateParam_Malilbox[iUnitId]:= TRUE;
aiTime1[iUnitId]:= aiTime1[iUnitId]+1;
					SysMemCpy(ADR(astStParam_Mailbox_out[iUnitId]),
							pstStParam_Mailbox_Tmp,
							SIZEOF(astStParam_Mailbox_out[iUnitId]));

					diTMP:= DWORD_TO_DINT(pstStParam_Mailbox_Tmp^.dwPlateAdjustmentProf);
					iUnitId_Tmp:= DWORD_TO_INT(DINT_TO_DWORD(diTMP) AND DWORD#255);(* 色组id *)
					diValue_Tmp:= SHR(diTMP, 8);(* 提交的数据 *)

					iRtn:=	KS_PushRapidAdjValue_V(ADR(g_astStAxisRapidAdjProf_V), iUnitId_Tmp, diValue_Tmp);
					IF iRtn <> 0 THEN
						(*2023.3.31.100107写日志2023.3.31.100110
						IF i_xRunlogEnable AND(* 2021.12.30.151304/日志使能 *)
							KS_IsValidUnitNR(iUnitId_Tmp) THEN
							sMsg_:= CONCAT('#SEMA_UPLOAD|KS_PushRapidAdjValue_V(Uid=', INT_TO_STRING(iUnitId_Tmp));
							sMsg_:= CONCAT(sMsg_, ')');
							KS_ThrowMsg2TravelLog(
								i_pstStTravelLogRec,
								LOG_LEVEL_INFO_DBG,
								sMsg_,
								DINT_TO_STRING(diValue_Tmp));
						END_IF
						*)
					ELSE
						;
					END_IF
IF pstStParam_Mailbox_Tmp^.iRapidAdjProf_h<>0 THEN
					(* 横向快速对版量 *)
					iRtn := KS_PushRapidAdjValue_H(ADR(g_astStAxisRapidAdjProf_H), iUnitId, pstStParam_Mailbox_Tmp^.iRapidAdjProf_h);

					IF iRtn <> 0 THEN
						(*2023.3.31.100107写日志2023.3.31.100110
						IF i_xRunlogEnable AND(* 2021.12.30.151345/日志使能 *)
							KS_IsValidUnitNR(iUnitNR) AND
							pstStProtocol_Mailbox_Tmp^.iRapidAdjProf_h<>0 THEN
							sMsg_:= CONCAT('#SEMA_UPLOAD|KS_PushRapidAdjValue_H(Uid=', INT_TO_STRING(iUnitNR));
							sMsg_:= CONCAT(sMsg_, ')');
							KS_ThrowMsg2TravelLog(
								i_pstStTravelLogRec,
								LOG_LEVEL_INFO_DBG,
								sMsg_,
								INT_TO_STRING(pstStProtocol_Mailbox_Tmp^.iRapidAdjProf_h));
						END_IF
						*)
					ELSE
						;
					END_IF
END_IF
					IF pastStParam_Mailbox_proof<>0 THEN(* 留存证据/下次比对用 *)
						SysMemCpy(ADR(pastStParam_Mailbox_proof^[iUnitId]), pstStParam_Mailbox_Tmp, SIZEOF(pstStParam_Mailbox_Tmp^));
					END_IF

					(* 正常接收的内容/就重新复位向量即可 *)
					pdwSEMA:= ADR(abyBuf_MailboxPkg_snd);
					IF pdwSEMA<>0 THEN
						pdwSEMA^:= SEMA_STANDBY;
//						iRtn:= GT_RN_DeviceLocalPcRamWr(pdwSEMA, DWORD_TO_WORD(dwOFST), KS_GetNumOfDwordUsed(SIZEOF(pdwSEMA^)));
						//SysMemCpy(ADR(abyBuf_MailboxPkg_snd), 1, SIZEOF(stStParam_Mailbox_Tmp));//2025.08.19 | TEST_
						iRtn:= GTN_RN_DevicePcMailWr(
								1,1,
								0,
								pdwSEMA,
								DWORD_TO_WORD(dwOFST),
								KS_GetNumOfDwordUsed(SIZEOF(pdwSEMA^)),
								16#1,0
								);

					END_IF
				ELSE
					(* 从站的参数非法/主动同步给从站/2021.12.4.142033/hdp *)
					SysMemCpy(ADR(stStParam_Mailbox_Tmp),ADR(astStParam_Mailbox_snd[iUnitId]),SIZEOF(stStParam_Mailbox_Tmp));
					//iRtn:= KS_FillUnitMailboxCmd_DN(ADR(stStParam_Mailbox_Tmp), pstStUnitParam_Save,pstStUnitParam_UnSave);
					SysMemSet(ADR(abyBuf_MailboxPkg_snd), 0, SIZEOF(abyBuf_MailboxPkg_snd));
					SysMemCpy(ADR(abyBuf_MailboxPkg_snd), ADR(stStParam_Mailbox_Tmp), SIZEOF(stStParam_Mailbox_Tmp));
//					iRtn:= GT_RN_DeviceLocalPcRamWr(ADR(abyBuf_MailboxPkg_snd), DWORD_TO_WORD(dwOFST), KS_GetNumOfDwordUsed(SIZEOF(pstStParam_Mailbox_Tmp)));
					//SysMemCpy(ADR(abyBuf_MailboxPkg_snd), 1, SIZEOF(stStParam_Mailbox_Tmp));//2025.08.19 | TEST_
					iRtn:= GTN_RN_DevicePcMailWr(
							1,1,
							0,
							ADR(abyBuf_MailboxPkg_snd),
							DWORD_TO_WORD(dwOFST),
							KS_GetNumOfDwordUsed(SIZEOF(pstStParam_Mailbox_Tmp)),
							16#1,0
							);
					IF iRtn<>0 THEN
						(*IF i_xRunlogEnable THEN(* 2021.12.21.133247/hdp *)
							KS_ThrowMsg2TravelLog(
								g_pstStTravelLogRec,
								LOG_LEVEL_INFO_DBG,
								'#SEMA_UPLOAD|Failed downloading...',
								INT_TO_STRING(iRtn));
						END_IF
						*);
					ELSE
						IF pastStParam_Mailbox_proof<>0 THEN(* 更新证据 *)
							(* 2023.11.22.093131/han.dp/已经修正过src地址和大小 *)
							SysMemCpy(ADR(pastStParam_Mailbox_proof^[iUnitId]), ADR(stStParam_Mailbox_Tmp), SIZEOF(stStParam_Mailbox_Tmp));
						END_IF
					END_IF

				END_IF

				(* 只要是约定的状态之一/就更新Mailbox通讯的超时时间/2021.12.21.135901/hdp *)
				atmUnitMailboxLastSynchronized[iUnitId]:= tmCURR;

			SEMA_DOWNLOAD:(* 主站下发的/从站还没有读取/要不再等等 *)
				(* 如果从站长时间不读取/本地数据又更新了/我们是不是考虑也把发送的内容更新一下 *)
				;

				(* 只要是约定的状态之一/就更新Mailbox通讯的超时时间/2021.12.21.135901/hdp *)
				atmUnitMailboxLastSynchronized[iUnitId]:= tmCURR;

			SEMA_PLS_REQ_DISPATCH:(* 请从站主动来请求 *)
				(* 等从站修改状态 *)
				;

				(* 只要是约定的状态之一/就更新Mailbox通讯的超时时间/2021.12.21.135901/hdp *)
				atmUnitMailboxLastSynchronized[iUnitId]:= tmCURR;

			SEMA_REQ_DISPATCH:(* 从站已经来请求了 *)
				(* 从站的参数非法/主动同步给从站/2021.12.4.142033/hdp *)
				SysMemCpy(ADR(stStParam_Mailbox_Tmp),ADR(astStParam_Mailbox_snd[iUnitId]),SIZEOF(stStParam_Mailbox_Tmp));

			//	iRtn:= KS_FillUnitMailboxCmd_DN(ADR(stStParam_Mailbox_Tmp), pstStUnitParam_Save,pstStUnitParam_UnSave);

				SysMemSet(ADR(abyBuf_MailboxPkg_snd), 0, SIZEOF(abyBuf_MailboxPkg_snd));
				SysMemCpy(ADR(abyBuf_MailboxPkg_snd), ADR(stStParam_Mailbox_Tmp), SIZEOF(stStParam_Mailbox_Tmp));

				//iRtn:= GT_RN_DeviceLocalPcRamWr(ADR(abyBuf_MailboxPkg_snd),
				//								DWORD_TO_WORD(dwOFST),
				//								KS_GetNumOfDwordUsed(SIZEOF(abyBuf_MailboxPkg_snd)));
				//改为实际长度2023.12.26.163451
// 				iRtn:= GTN_RN_DeviceLocalPcRamWr(ADR(abyBuf_MailboxPkg_snd),
// 												DWORD_TO_WORD(dwOFST),
// 												KS_GetNumOfDwordUsed(SIZEOF(stStParam_Mailbox_Tmp)));
				iRtn:= GTN_RN_DevicePcMailWr(
						1,1,
						0,
						ADR(abyBuf_MailboxPkg_snd),
						DWORD_TO_WORD(dwOFST),
						KS_GetNumOfDwordUsed(SIZEOF(stStParam_Mailbox_Tmp)),
						16#1,0
						);
(*
FUNCTION GTN_RN_DevicePcMailWr : INT
VAR_INPUT
	cardIndex:INT;
	busIndex:INT;
	stationId:INT;
	pData:POINTER TO UDINT;
	startAddr:UINT;
	dwordNum:UINT;
	cmdType:BYTE;
	respReq:BYTE;
END_VAR
VAR
END_VAR
*)

				IF iRtn<>0 THEN
					(*IF i_xRunlogEnable THEN(* 2021.12.21.132943/hdp *)
						KS_ThrowMsg2TravelLog(
							g_pstStTravelLogRec,
							LOG_LEVEL_INFO_DBG,
							'#SEMA_REQ_DISPATCH|Failed downloading...',
							INT_TO_STRING(iRtn));
					END_IF
					*);
				ELSE
					IF pastStParam_Mailbox_proof<>0 THEN(* 更新证据 *)
						(* 2023.11.22.093131/han.dp/已经修正过src地址和大小 *)
						SysMemCpy(ADR(pastStParam_Mailbox_proof^[iUnitId]), ADR(stStParam_Mailbox_Tmp), SIZEOF(stStParam_Mailbox_Tmp));
					END_IF
				END_IF

				(* 只要是约定的状态之一/就更新Mailbox通讯的超时时间/2021.12.21.135901/hdp *)
				atmUnitMailboxLastSynchronized[iUnitId]:= tmCURR;
			ELSE
				(* 剩余的情况/就定期扫描看主站数据是否有更新 *)
				(* 定期强行同步的机制取消掉/改为从站60s(暂定)没有收到主站的数据/主动发送SEMA_REQ_DISPATCH信号过来要参数 *)
				IF pastStParam_Mailbox_proof<>0 THEN(* 证据可以访问 *)

					pdata1:= ADR(astStParam_Mailbox_snd[iUnitId]);
					pdata2:= ADR(pastStParam_Mailbox_proof^[iUnitId]);

					pdata1:= pdata1+4;
					pdata2:= pdata2+4;
					xFlag_MasterChange:= FALSE;
					iLength:= SIZEOF(astStParam_Mailbox_snd[iUnitId])-4;
					FOR iK:=1 TO iLength BY 1 DO
						IF pdata1^<>pdata2^ THEN
							xFlag_MasterChange:=TRUE;
							EXIT;
						END_IF
						pdata1:= pdata1+1;
						pdata2:= pdata2+1;
					END_FOR
					IF 	xFlag_MasterChange THEN
						SysMemCpy(ADR(stStParam_Mailbox_Tmp),ADR(astStParam_Mailbox_snd[iUnitId]),SIZEOF(stStParam_Mailbox_Tmp));
					//	iRtn:= KS_FillUnitMailboxCmd_DN(ADR(stStParam_Mailbox_Tmp), pstStUnitParam_Save,pstStUnitParam_UnSave);

						SysMemSet(ADR(abyBuf_MailboxPkg_snd), 0, SIZEOF(abyBuf_MailboxPkg_snd));
						SysMemCpy(ADR(abyBuf_MailboxPkg_snd), ADR(stStParam_Mailbox_Tmp), SIZEOF(stStParam_Mailbox_Tmp));

						//SysMemCpy(ADR(abyBuf_MailboxPkg_snd), 1, SIZEOF(stStParam_Mailbox_Tmp));//2025.08.19 | TEST_
						iRtn:= GTN_RN_DevicePcMailWr(
									1,1,0,
									ADR(abyBuf_MailboxPkg_snd),
									DWORD_TO_WORD(dwOFST),
									KS_GetNumOfDwordUsed(SIZEOF(stStParam_Mailbox_Tmp)),
									RN_AWR,
									0);
						IF iRtn<>0 THEN
							(*IF i_xRunlogEnable THEN(* 2021.12.21.132817/hdp *)
								KS_ThrowMsg2TravelLog(
									g_pstStTravelLogRec,
									LOG_LEVEL_INFO_DBG,
									'#ELSE|Failed downloading...',
									INT_TO_STRING(iRtn));
							END_IF
							*);
						ELSE
							IF pastStParam_Mailbox_proof<>0 THEN(* 更新证据 *)
								SysMemCpy(ADR(pastStParam_Mailbox_proof^[iUnitId]), ADR(stStParam_Mailbox_Tmp), SIZEOF(stStParam_Mailbox_Tmp));
							END_IF
						END_IF

						(* 只要是约定的状态之一/就更新Mailbox通讯的超时时间/2021.12.21.135901/hdp *)
						atmUnitMailboxLastSynchronized[iUnitId]:= tmCURR;

					ELSE(* 主站的参数一直没发生修改/超过3s从站不响应/就让从站重新请求 *)
						IF tmCURR-atmUnitMailboxLastSynchronized[iUnitId]>=TIMEOUTS_MAILBOX_FORCESYNC THEN
							pdwSEMA:= ADR(abyBuf_MailboxPkg_snd);
							IF pdwSEMA<>0 THEN
								pdwSEMA^:= SEMA_PLS_REQ_DISPATCH;
								//SysMemCpy(ADR(abyBuf_MailboxPkg_snd), 1, SIZEOF(stStParam_Mailbox_Tmp));//2025.08.19 | TEST_
								iRtn:= GTN_RN_DevicePcMailWr(
										1,1,0,
										pdwSEMA,
										DWORD_TO_WORD(dwOFST),
										KS_GetNumOfDwordUsed(SIZEOF(pdwSEMA^)),
										RN_AWR,
										0);
							END_IF

							(* 只要是约定的状态之一/就更新Mailbox通讯的超时时间/2021.12.21.135901/hdp *)
							atmUnitMailboxLastSynchronized[iUnitId]:= tmCURR;
						END_IF
					END_IF
				ELSE
					(* 作为存档的参考内存无法申请到/pastStProtocol_Mailbox_proof *)
					(*IF i_xRunlogEnable THEN(* 2021.12.21.133109/hdp *)
						KS_ThrowMsg2TravelLog(
							g_pstStTravelLogRec,
							LOG_LEVEL_INFO_DBG,
							'#BAD POINTER',
							'pastStProtocol_Mailbox_proof');
					END_IF
					*);
				END_IF
			END_CASE
		ELSE
			;
		END_IF
	ELSE
		;
	END_IF
END_FOR

(* ---- Action_RdSampleData.st ---- *)
(*@CES
Name=Action_RdSampleData
Type=Action
TypeGuid=8ac092e5-3128-4e26-9e7e-11016c6684f2
Guid=9712102a-3aaf-4685-ba49-06f5bfb943ae
HasDeclaration=False
HasImplementation=True
*)
{DECLARATION}

{IMPLEMENTATION}

iUMax_Tmp:= g_stStSysParam.stStSysParam_Save.iUnitMaxNum;
iUid_Tmp:= g_stStSysParam.stStSysParam_Save.iUid;
IF iUid_Tmp>=2 AND iUid_Tmp<= iUMax_Tmp THEN
	IF NOT g_stStSysParam.astStUnitParam_Save[iUid_Tmp].xEnable_arc THEN
		xReDirectedCurrUnit:= TRUE;
	END_IF
ELSE
	xReDirectedCurrUnit:= TRUE;
END_IF

IF xReDirectedCurrUnit THEN(*需要重新定向|找第1个使能套色的色组|*)
	FOR iN:=2 TO iUMax_Tmp BY 1 DO
		IF g_stStSysParam.astStUnitParam_Save[iN].xEnable_arc THEN
			g_stStSysParam.stStSysParam_Save.iUid := iN;
			xReDirectedCurrUnit := FALSE;//2025.11.19.151125 | 重定向完成
			EXIT;
		END_IF
	END_FOR
END_IF
IF g_stStSysParam.stStSysParam_Save.iUid<> iLastId AND
		g_stStSysParam.stStSysParam_Save.iUid>=2 AND
		g_stStSysParam.stStSysParam_Save.iUid<=g_stStSysParam.stStSysParam_Save.iUnitMaxNum THEN
	iLastId:= g_stStSysParam.stStSysParam_Save.iUid;
	iStationId:= g_stStSysParam.stStSysParam_UnSave.aiStationList_UnitController[g_stStSysParam.stStSysParam_Save.iUid];
	IF iStationId<>-1 THEN
		aiRtnCode[1]:= GT_RN_SampleSetShowDeviceId(INT_TO_BYTE(iStationId));
		aiRtnCode[2]:= GT_RN_SampleRoundUpdata();
	END_IF
END_IF
(*
byChannael-bit0:T2-R
		   bit1:T2-G
		   bit2:T2-B
		   bit4:T1-R
		   bit5:T1-G
		   bit6:T1-B
*)
aiRtnCode[3]:= GT_RN_SampleGetRoundDataEx(
					g_stStSysParam.astStUnitParam_Save[g_stStSysParam.stStSysParam_Save.iUid].bySignalSelect,
					ADR(g_pbyRoundData1),
					ADR(g_pbyRoundData2),
					ADR(iRoundSampleFlag));

IF iRoundSampleFlag=1 THEN
	IF g_pbyRoundData2<>0 AND g_pbyRoundData1<>0 THEN
		IF g_stStSysParam.astStUnitParam_Save[g_stStSysParam.stStSysParam_Save.iUid].bySignalSelect.0 THEN
			SysMemCpy(ADR(g_stStSysParam.stStSysParam_UnSave.abyData_T1_R),
						g_pbyRoundData1,
						SIZEOF(g_stStSysParam.stStSysParam_UnSave.abyData_T1_R));

		ELSIF g_stStSysParam.astStUnitParam_Save[g_stStSysParam.stStSysParam_Save.iUid].bySignalSelect.1 THEN
			SysMemCpy(ADR(g_stStSysParam.stStSysParam_UnSave.abyData_T1_G),
						g_pbyRoundData1,
						SIZEOF(g_stStSysParam.stStSysParam_UnSave.abyData_T1_G));

		ELSIF g_stStSysParam.astStUnitParam_Save[g_stStSysParam.stStSysParam_Save.iUid].bySignalSelect.2 THEN
			SysMemCpy(ADR(g_stStSysParam.stStSysParam_UnSave.abyData_T1_B),
						g_pbyRoundData1,
						SIZEOF(g_stStSysParam.stStSysParam_UnSave.abyData_T1_B));
		ELSE
			SysMemCpy(ADR(g_stStSysParam.stStSysParam_UnSave.abyData_T1_R),
						g_pbyRoundData1,
						SIZEOF(g_stStSysParam.stStSysParam_UnSave.abyData_T1_R));
		END_IF
		IF g_stStSysParam.astStUnitParam_Save[g_stStSysParam.stStSysParam_Save.iUid].bySignalSelect.4 THEN
			SysMemCpy(ADR(g_stStSysParam.stStSysParam_UnSave.abyData_T2_R),
						g_pbyRoundData2,
						SIZEOF(g_stStSysParam.stStSysParam_UnSave.abyData_T2_R));
		ELSIF g_stStSysParam.astStUnitParam_Save[g_stStSysParam.stStSysParam_Save.iUid].bySignalSelect.5 THEN
			SysMemCpy(ADR(g_stStSysParam.stStSysParam_UnSave.abyData_T2_G),
						g_pbyRoundData2,
						SIZEOF(g_stStSysParam.stStSysParam_UnSave.abyData_T2_G));
		ELSIF g_stStSysParam.astStUnitParam_Save[g_stStSysParam.stStSysParam_Save.iUid].bySignalSelect.6 THEN
			SysMemCpy(ADR(g_stStSysParam.stStSysParam_UnSave.abyData_T2_B),
						g_pbyRoundData2,
						SIZEOF(g_stStSysParam.stStSysParam_UnSave.abyData_T2_B));
		ELSE
			SysMemCpy(ADR(g_stStSysParam.stStSysParam_UnSave.abyData_T2_R),
						g_pbyRoundData2,
						SIZEOF(g_stStSysParam.stStSysParam_UnSave.abyData_T2_R));
		END_IF
		(*2026.5.9.144620*)
		(*2026.03.23.171805||保存采样wang.xy*)
		IF g_stStSysParam.stStSysParam_Save.iUid>=2 AND
			g_stStSysParam.stStSysParam_Save.iUid<=g_stStSysParam.stStSysParam_Save.iUnitMaxNum THEN
			KS_PshRSdata2Fifo(
				g_pstStRSampFifo,
				g_pbyRoundData1,
				g_pbyRoundData2,
				INT_TO_BYTE(g_stStSysParam.stStSysParam_Save.iUid),
				LREAL_TO_DINT(g_stStSysParam.astStUnitParam_UnSave[g_stStSysParam.stStSysParam_Save.iUid].rAxisVel_PrnRoller*100.0),
				g_astStTaskCycleDetection[1].udiCycleCnt);
		END_IF

	END_IF
	aiRtnCode[4]:= GT_RN_SampleRoundUpdata();(* 启动下一次采样 *)
ELSE
		(*2026.03.23.162723||粗采样保存wang.xy*)
	fbKS_FB_ExportRSFifo2File(
//		i_xEn:= g_xSaveRS2file,2026.5.14.091655更新屏蔽
		i_xEn:= g_stStSysParam.astStRSV_GrpParam_UnSave[1].xSwitch_SaveRS2file,
		i_sPath:= ,
		i_pstStRSampFifo:= g_pstStRSampFifo,
		o_iErNo=> iRtn);
END_IF

(* ---- Action_SyncParamToSample.st ---- *)
(*@CES
Name=Action_SyncParamToSample
Type=Action
TypeGuid=8ac092e5-3128-4e26-9e7e-11016c6684f2
Guid=a15681d5-bd2f-4cd2-a15c-8116b58af265
HasDeclaration=False
HasImplementation=True
*)
{DECLARATION}

{IMPLEMENTATION}
(* 首次同步参数记录|用以后续检查变动了没有|@2018.5.21.095735 *)
IF NOT xSynchronized_SpecialParam THEN
	xSynchronized_SpecialParam:= TRUE;
	FOR iGrp:=1 TO 2 BY 1 DO
		aiMarkTypeId[iGrp]:= g_stStSysParam.astStGrpParam_Save[iGrp].iMarkTypeId;
		aiMarkArrangeId[iGrp]:= g_stStSysParam.astStGrpParam_Save[iGrp].iMarkArrangeMode;
	END_FOR
END_IF

FOR iGrp:=1 TO 2 BY 1 DO

(* 同步系内的全局设定到色组同步|@2017.8.3.085112 *)
	pstStGrpParam_Save:= ADR(g_stStSysParam.astStGrpParam_Save[iGrp]);
	pstStGrpParam_UnSave:= ADR(g_stStSysParam.astStGrpParam_UnSave[iGrp]);

	(* 标记形式 *)
	IF aiMarkTypeId[iGrp]<>pstStGrpParam_Save^.iMarkTypeId THEN
		FOR iN:=1 TO MAX_UNIT_NUM BY 1 DO
			pstStUnitParam_Save:= ADR(g_stStSysParam.astStUnitParam_Save[iN]);
			pstStUnitParam_UnSave:= ADR(g_stStSysParam.astStUnitParam_UnSave[iN]);

			IF pstStUnitParam_Save^.byGrpId=INT_TO_BYTE(iGrp) THEN
				pstStUnitParam_Save^.iMarkTypeId:= pstStGrpParam_Save^.iMarkTypeId;
			END_IF

		END_FOR
		aiMarkTypeId[iGrp]:= pstStGrpParam_Save^.iMarkTypeId;
	END_IF

(*2025.9.20.103056这里处理放到金刚吧
	(* 标记排列|当选择横排和纵排切换的时候|需要把门内基线自动切换一下|@2019.11.14.102415 *)
	IF aiMarkArrangeId[iGrp]<>pstStGrpParam_Save^.iMarkArrangeMode THEN
		FOR iN:=1 TO MAX_UNIT_NUM BY 1 DO
			pstStUnitParam_Save:= ADR(g_stStSysParam.astStUnitParam_Save[iN]);
			pstStUnitParam_UnSave:= ADR(g_stStSysParam.astStUnitParam_UnSave[iN]);
			IF pstStUnitParam_Save^.byGrpId=INT_TO_BYTE(iGrp) THEN
				pstStUnitParam_Save^.iMarkArrangeMode:= pstStGrpParam_Save^.iMarkArrangeMode;
				CASE pstStUnitParam_Save^.iMarkArrangeMode OF
				MARK_ARRANGE_HFOR,MARK_ARRANGE_HREV:(*横排|*)
					IF NOT (aiMarkArrangeId[iGrp]=MARK_ARRANGE_HFOR OR aiMarkArrangeId[iGrp]=MARK_ARRANGE_HREV) THEN
						(* 如果之前是纵排 *)
						IF NOT pstStUnitParam_Save^.dwFlag_Ctl.1 THEN (* 如果没打开门内基线|则我们帮助其默认打开 *)
							pstStUnitParam_Save^.dwFlag_Ctl.1:= TRUE;
						END_IF
					END_IF
				ELSE(*全部当纵排处理|*)
					IF aiMarkArrangeId[iGrp]=MARK_ARRANGE_HFOR OR aiMarkArrangeId[iGrp]=MARK_ARRANGE_HREV THEN
						(* 如果之前是横排 *)
						IF pstStUnitParam_Save^.dwFlag_Ctl.1 THEN (* 如果打开了门内基线|则我们帮助其默认关闭 *)
							pstStUnitParam_Save^.dwFlag_Ctl.1:= FALSE;
						END_IF
					END_IF
				END_CASE
			END_IF
		END_FOR
		aiMarkArrangeId[iGrp]:= pstStGrpParam_Save^.iMarkArrangeMode;(*移动到最后更新|2019.11.14.103051_*)
	END_IF
	*)
END_FOR

FOR iN:=1 TO g_stStSysParam.stStSysParam_Save.iUnitMaxNum(*g_pstStShmGlobalParam^.iUMax*) BY 1 DO
	(* 条标时把横向打开了|系统强制关闭|@2019.4.26.133820 *)
	IF g_stStSysParam.astStUnitParam_Save[iN].iMarkTypeId=MARK_TYPE_LINE AND
		g_stStSysParam.astStUnitParam_Save[iN].dwFlag_Ctl.0 THEN
		g_stStSysParam.astStUnitParam_Save[iN].dwFlag_Ctl.0:= FALSE; (* 关横向 *)
	END_IF

	(*横向手动版修正|*)
	IF NOT axSynchronizedFlag[iN] THEN
		axSynchronizedFlag[iN]:= TRUE;
	ELSE
		IF g_abyHorzManu_HMI[iN].0<>abyHorzManu_HMI_Pre[iN].0 THEN (* 横向左手动1 *)
			g_abyHorzManuTrigButton[iN]:= 1;
			KS_HY_AddMsgToLog(g_pstStHYLogFifo,
				LOG_LEVEL_EVT_USRACTIONS, 'Horz-Manu-Adj-Left-1', INT_TO_STRING(iN)); (* 2020.8.11.141918|watching... *)
		END_IF
		IF g_abyHorzManu_HMI[iN].1<>abyHorzManu_HMI_Pre[iN].1 THEN (* 横向左手动2 *)
			g_abyHorzManuTrigButton[iN]:= 2;
			KS_HY_AddMsgToLog(g_pstStHYLogFifo,
				LOG_LEVEL_EVT_USRACTIONS, 'Horz-Manu-Adj-Left-2', INT_TO_STRING(iN)); (* 2020.8.11.141918|watching... *)
		END_IF
		IF g_abyHorzManu_HMI[iN].2<>abyHorzManu_HMI_Pre[iN].2 THEN (* 横向右手动1 *)
			g_abyHorzManuTrigButton[iN]:= 3;
			KS_HY_AddMsgToLog(g_pstStHYLogFifo,
				LOG_LEVEL_EVT_USRACTIONS, 'Horz-Manu-Adj-Right-1', INT_TO_STRING(iN)); (* 2020.8.11.141918|watching... *)
		END_IF
		IF g_abyHorzManu_HMI[iN].3<>abyHorzManu_HMI_Pre[iN].3 THEN (* 横向右手动2 *)
			g_abyHorzManuTrigButton[iN]:= 4;
			KS_HY_AddMsgToLog(g_pstStHYLogFifo,
				LOG_LEVEL_EVT_USRACTIONS, 'Horz-Manu-Adj-Right-2', INT_TO_STRING(iN)); (* 2020.8.11.141918|watching... *)
		END_IF

(*2022.8.9.092113||更新韩工7.29更新||横向手动按钮0.02档位*)
		IF g_abyHorzManu_HMI[iN].4<>abyHorzManu_HMI_Pre[iN].4 THEN (* 横向左0.02 *)
			g_abyHorzManuTrigButton[iN]:= 5;
			KS_HY_AddMsgToLog(g_pstStHYLogFifo,
				LOG_LEVEL_EVT_USRACTIONS, 'Horz-Manu-Adj-Left-3', INT_TO_STRING(iN)); (* 2020.8.11.141918|watching... *)
		END_IF

		IF g_abyHorzManu_HMI[iN].5<>abyHorzManu_HMI_Pre[iN].5 THEN (* 横向右0.02 *)
			g_abyHorzManuTrigButton[iN]:= 6;
			KS_HY_AddMsgToLog(g_pstStHYLogFifo,
				LOG_LEVEL_EVT_USRACTIONS, 'Horz-Manu-Adj-Right-3', INT_TO_STRING(iN)); (* 2020.8.11.141918|watching... *)
		END_IF

	END_IF
	abyHorzManu_HMI_Pre[iN]:= g_abyHorzManu_HMI[iN];

END_FOR

wAxis_RollerDn:= 0;
wAxis_Alarm_Prn:= 0;
dwAlarmCode:= 0;
wComplexFlag_AxisInching:= 0;
wComplexFlag_Linkage:= 0;
wComplexFlag_Estop:= 0;

FOR iN:=1 TO MAX_UNIT_NUM BY 1 DO
	IF g_stStSysParam.astStUnitParam_Save[iN].xLinkage THEN
		wComplexFlag_Linkage:= wComplexFlag_Linkage OR SHL(WORD#1, iN-1);
	END_IF

	IF g_stStSysParam.astStUnitParam_UnSave[iN].xAxisInching OR g_axAxisInchDecing[iN] THEN
		wComplexFlag_AxisInching:= wComplexFlag_AxisInching OR SHL(WORD#1, iN-1);
	END_IF
	IF g_astStIOMap_Axis_FE[iN].o_xRel_Press THEN
		wAxis_RollerDn:= wAxis_RollerDn OR SHL(WORD#1, iN-1);
	END_IF
END_FOR

(* ---- Action_Udp_UnitHMI.st ---- *)
(*@CES
Name=Action_Udp_UnitHMI
Type=Action
TypeGuid=8ac092e5-3128-4e26-9e7e-11016c6684f2
Guid=cdb6e806-737e-4889-9ab9-78f8b741b17a
HasDeclaration=False
HasImplementation=True
*)
{DECLARATION}

{IMPLEMENTATION}
(*2025.6.23.144921|niu.j||子影人机通讯*)
(*先获取上次通讯的响应码*)
IF NOT xInit_Comm_HMI THEN
	xInit_Comm_HMI:= TRUE;
	(*初始化*)
	FOR iN:=1 TO MAX_UNIT_NUM BY 1 DO
		iUnitId:= iN;
		axFlag_Comm_ReadEn[iUnitId] := FALSE;
		(*初始化网络*)
		aiStep_Comm[iUnitId]:= 3;
	END_FOR
	iUnitId_To_Hmi:= 1;
	//g_abyStationList_CommHMI;
END_IF

IF iUnitId_To_Hmi>g_stStSysParam.stStSysParam_Save.iUnitMaxNum THEN(*只需要循环到最大色组*)
	iUnitId_To_Hmi:= 1;
END_IF
iUnitId:= iUnitId_To_Hmi;
SysMemSet(ADR(abyBuf_UDP_Unit_rcv[iUnitId,1]),0,MAILBOX_PKG_MAX_BYTES);

(*先同步一次参数后再开始读取响应*)
// 	iUnitNR:=1;
// 	dwOFST:= INT_TO_DWORD((iUnitNR-1))*MAILBOX_PKG_MAX_BYTES;
dwOFST:= INT_TO_DWORD((iUnitId-1))*INT_TO_DWORD(MAILBOX_PKG_MAX_BYTES);
(*iStationId:= g_abyStationList_CommHMI[iN];*)
iStationId:= g_abyStationList_CommHMI[iUnitId];

SysMemSet(ADR(abyBuf_UDP_Unit_rcv_Use_Tmp[iUnitId]),0,SIZEOF(abyBuf_UDP_Unit_rcv_Use_Tmp[iUnitId]));
IF KS_IsValidStationNR(iStationId) AND KS_IsValidUnitNR(iUnitId) THEN
	(*GTN_RN_DevicePcMailRd(
		1,2,
		0,
		ADR(abyBuf_UDP_Unit_rcv[iUnitId,1]),
		DWORD_TO_UINT(dwOFST),
		KS_GetNumOfDwordUsed(MAILBOX_PKG_MAX_BYTES),
		RN_ARD
		);*)
	IF g_abyStationList_CommHMI[iUnitId]<=0 THEN
		iUnitId_To_Hmi:= iUnitId_To_Hmi+1;
		RETURN;
	END_IF
	iRtn1:=GTN_RN_DevicePcMailRd(
		1,2,
		iStationId,
		ADR(abyBuf_UDP_Unit_rcv[iUnitId,1]),
		0,//DWORD_TO_UINT(dwOFST),
		KS_GetNumOfDwordUsed(MAILBOX_PKG_MAX_BYTES),
		RN_ARD
		);
	IF aiStep_Comm[iUnitId]>2 THEN
		axFlag_DataCmd[iUnitId]:=TRUE;
	ELSE
		IF abyBuf_UDP_Unit_snd[iUnitId,2]= SEMA_FUNCODE_485_MULT_RD THEN
			axFlag_DataCmd[iUnitId]:=FALSE;
		ELSE
			axFlag_DataCmd[iUnitId]:=TRUE;
		END_IF
	END_IF
	//abyRdDataNum[iUnitId]:=word_to_byte(KS_GetNumOfDwordUsed(MAILBOX_PKG_MAX_BYTES));
	KS_Modbus_ReadFun(
		TRUE,(*i_xEn:= , *)
		1,(*i_byType_RegisterorCoils:= , *)
		axFlag_DataCmd[iUnitId],(*i_xFlag_DataCmd:= , *)
		iUnitId,(*i_iUnitId_Tar:= , *)
		abyRdDataNum[iUnitId],(*i_byRdDataNum:= , *)
		ADR(abyBuf_UDP_Unit_rcv[iUnitId,1]),(*i_pbyDataBf:= , *)
		ADR(abyBuf_UDP_Unit_rcv_Use_Tmp)(*i_pbyDataRd_Use:= *));
	(*根据收到的响应内容，-处理有效数据*)
	IF axFlag_Rd_OR_WrRd[iUnitId] THEN
		SysMemCpy(ADR(astStParam_UnitHMI485_WrRd[iUnitId]),//收到的数据
			ADR(abyBuf_UDP_Unit_rcv_Use_Tmp),
			SIZEOF(astStParam_UnitHMI485_WrRd[iUnitId]));
		SysMemCpy(ADR(astStParam_UnitHMI485_WrRd_Rec[iUnitId]),
			ADR(astStParam_UnitHMI485_WrRd[iUnitId]),
			SIZEOF(astStParam_UnitHMI485_WrRd_Rec[iUnitId]));
		axFlag_Rd_Or_WrRd[iUnitId]:= FALSE;
	ELSE
		SysMemCpy(ADR(astStParam_UnitHMI485_Rd[iUnitId]),
			ADR(abyBuf_UDP_Unit_rcv_Use_Tmp),
			SIZEOF(astStParam_UnitHMI485_Rd[iUnitId]));
	END_IF
	aiStep_Comm[iUnitId]:= aiStep_Comm[iUnitId]+1;
	IF aiStep_Comm[iUnitId]>5 THEN
		aiStep_Comm[iUnitId]:=1;
	END_IF
	(*响应码处理完成-处理写入数据*)
	(*先判断读写参数有没有变化*)
	diTemp:= 0;
	astStParam_UnitHMI485_WrRd[iUnitId].byAxisId:= INT_TO_BYTE(iUnitId);
	diTemp:=DWORD_TO_DINT(SysMemCmp(ADR(astStParam_UnitHMI485_WrRd_Rec[iUnitId]),
			ADR(astStParam_UnitHMI485_WrRd[iUnitId]),
			SIZEOF(astStParam_UnitHMI485_WrRd_Rec[iUnitId])));
	SysMemCpy(ADR(astStParam_UnitHMI485_WrRd_Rec[iUnitId]),
		ADR(astStParam_UnitHMI485_WrRd[iUnitId]),
		SIZEOF(astStParam_UnitHMI485_WrRd_Rec[iUnitId]));
	IF diTemp=0 THEN
		CASE aiStep_Comm[iUnitId] OF
			(*写入数据流程-读-读-写-写*)
			1:
			KS_Modbus_WriteFun(
				TRUE,(*i_xEn:= , *)
				1,(*i_byType_RegisterorCoils:= , *)
				FALSE,(*i_xFlag_DataCmd:= , *)
				iUnitId,(*i_iUnitId_Tar:= , *)
				600,(*i_wAddr_Comm:= , *)(*双向数据的通讯地址*)
				ADR(astStParam_UnitHMI485_WrRd[iUnitId]),(*i_pData_Addrstart:= , *)
				240,(*i_byLength_Data:= *)
				ADR(abyBuf_UDP_Unit_snd[iUnitId,1]));
			abyRdDataNum[iUnitId]:= 245;
			axFlag_Rd_Or_WrRd[iUnitId]:= TRUE;
			2:
			KS_Modbus_WriteFun(
				TRUE,(*i_xEn:= , *)
				1,(*i_byType_RegisterorCoils:= , *)
				FALSE,(*i_xFlag_DataCmd:= , *)
				iUnitId,(*i_iUnitId_Tar:= , *)
				720,(*i_wAddr_Comm:= , *)(*双向数据的通讯地址*)
				ADR(astStParam_UnitHMI485_Rd[iUnitId]),(*i_pData_Addrstart:= , *)
				240,(*i_byLength_Data:= *)
				ADR(abyBuf_UDP_Unit_snd[iUnitId,1]));
			abyRdDataNum[iUnitId]:= 245;
			3:
			KS_Modbus_WriteFun(
				TRUE,(*i_xEn:= , *)
				1,(*i_byType_RegisterorCoils:= , *)
				TRUE,(*i_xFlag_DataCmd:= , *)
				iUnitId,(*i_iUnitId_Tar:= , *)
				0,(*i_wAddr_Comm:= , *)(*双向数据的通讯地址*)
				ADR(astStParam_UnitHMI485_Wr_81[iUnitId]),(*i_pData_Addrstart:= , *)
				240,(*i_byLength_Data:= *)
				ADR(abyBuf_UDP_Unit_snd[iUnitId,1]));
			abyRdDataNum[iUnitId]:= 8;
			4:
			KS_Modbus_WriteFun(
				TRUE,(*i_xEn:= , *)
				1,(*i_byType_RegisterorCoils:= , *)
				TRUE,(*i_xFlag_DataCmd:= , *)
				iUnitId,(*i_iUnitId_Tar:= , *)
				120,(*i_wAddr_Comm:= , *)(*双向数据的通讯地址*)
				ADR(astStParam_UnitHMI485_Wr_82[iUnitId]),(*i_pData_Addrstart:= , *)
				240,(*i_byLength_Data:= *)
				ADR(abyBuf_UDP_Unit_snd[iUnitId,1]));
			abyRdDataNum[iUnitId]:= 8;
			5:
			KS_Modbus_WriteFun(
				TRUE,(*i_xEn:= , *)
				1,(*i_byType_RegisterorCoils:= , *)
				TRUE,(*i_xFlag_DataCmd:= , *)
				iUnitId,(*i_iUnitId_Tar:= , *)
				360,(*i_wAddr_Comm:= , *)(*双向数据的通讯地址*)
				ADR(astStParam_UnitHMI485_Wr_83[iUnitId]),(*i_pData_Addrstart:= , *)
				240,(*i_byLength_Data:= *)
				ADR(abyBuf_UDP_Unit_snd[iUnitId,1]));
			abyRdDataNum[iUnitId]:= 8;
		END_CASE
	ELSE
		KS_Modbus_WriteFun(
			TRUE,(*i_xEn:= , *)
			1,(*i_byType_RegisterorCoils:= , *)
			TRUE,(*i_xFlag_DataCmd:= , *)
			iUnitId,(*i_iUnitId_Tar:= , *)
			600,(*i_wAddr_Comm:= , *)(*双向数据的通讯地址*)
			ADR(astStParam_UnitHMI485_WrRd[iUnitId]),(*i_pData_Addrstart:= , *)
			UINT_TO_BYTE(SIZEOF(astStParam_UnitHMI485_WrRd[iUnitId]))(*i_byLength_Data:= *),
			ADR(abyBuf_UDP_Unit_snd[iUnitId,1]));
		abyRdDataNum[iUnitId]:= 8;
	END_IF

	 iRtn2:=GTN_RN_DevicePcMailWr(
		1,2,
		iStationId,
		ADR(abyBuf_UDP_Unit_snd[iUnitId,1]),
		//abyBuf_UDP_Unit_snd[iUnitId,1],
		0,//DWORD_TO_UINT(dwOFST),
		KS_GetNumOfDwordUsed(MAILBOX_PKG_MAX_BYTES),
		RN_AWR,
		0
		);
END_IF
iUnitId_To_Hmi:= iUnitId_To_Hmi+1;(*循环下一个色组*)

(* ---- Action_Udp_UnitHMI_Input.st ---- *)
(*@CES
Name=Action_Udp_UnitHMI_Input
Type=Action
TypeGuid=8ac092e5-3128-4e26-9e7e-11016c6684f2
Guid=f5c1d7ba-7edb-4795-af5d-1ee2ef07b11e
HasDeclaration=False
HasImplementation=True
*)
{DECLARATION}

{IMPLEMENTATION}
FOR iN:=1 TO MAX_UNIT_NUM BY 1 DO
	iGrpIdTmp:= g_stStSysParam.astStUnitParam_Save[iN].byGrpId;
	astStParam_UnitHMI485_Wr_81[iN].byPackId:= 1;
	astStParam_UnitHMI485_Wr_81[iN].wGirth:= REAL_TO_WORD(g_stStSysParam.astStUnitParam_Save[iN].rGirth_Sam*10);
	astStParam_UnitHMI485_Wr_81[iN].iCompanyId:= g_stStSysParam.stStSysParam_Save.iCustomerId;
	astStParam_UnitHMI485_Wr_81[iN].iPromptMsgId:= g_stStSysParam.astStGrpParam_UnSave[iGrpIdTmp].iPromptMsg;
	astStParam_UnitHMI485_Wr_81[iN].wAxisId_And_GrpId:= SHL(INT_TO_WORD(iN),8)+INT_TO_WORD(iGrpIdTmp);
	astStParam_UnitHMI485_Wr_81[iN].wLedtime_And_Language:= SHL(BYTE_TO_WORD(g_stStSysParam.stStSysParam_Save.byMinutes_ScrSaver),8)+
																BYTE_TO_WORD(g_stStSysParam.stStSysParam_Save.byLanguageId);
	astStParam_UnitHMI485_Wr_81[iN].iVel_Axis:= REAL_TO_INT(g_stStSysParam.astStUnitParam_UnSave[iN].rAxisVel_PrnRoller*10.0);
	astStParam_UnitHMI485_Wr_81[iN].iVel_Grp:= REAL_TO_INT(g_stStSysParam.astStGrpParam_UnSave[iGrpIdTmp].rVel_Cur*10.0);
	astStParam_UnitHMI485_Wr_81[iN].wIndex_And_ErrNum:= g_stStSysParam.astStUnitParam_UnSave[iN].byIndex;
	astStParam_UnitHMI485_Wr_81[iN].iArcAlarm_V:= REAL_TO_INT(g_stStSysParam.astStUnitParam_Save[iN].rAlr_V*100);//单位丝
	astStParam_UnitHMI485_Wr_81[iN].iArcAlarm_H:= REAL_TO_INT(g_stStSysParam.astStUnitParam_Save[iN].rAlr_H*100);//单位丝
	astStParam_UnitHMI485_Wr_81[iN].wUnit_Input_I:= g_stStSysParam.astStUnitParam_UnSave[iN].wUnit_input_I;
	astStParam_UnitHMI485_Wr_81[iN].wUnit_Input_II:= g_stStSysParam.astStUnitParam_UnSave[iN].wUnit_input_II;
	astStParam_UnitHMI485_Wr_81[iN].wUnit_Input_III:= g_stStSysParam.astStUnitParam_UnSave[iN].wUnit_input_III;
	astStParam_UnitHMI485_Wr_81[iN].wHz_UnitInkRoller_CurrWR:= REAL_TO_WORD(g_stStSysParam.astStUnitParam_UnSave[iN].rHz_UnitInkRoller_CurrWR*100);
	astStParam_UnitHMI485_Wr_81[iN].wHz_UnitScraper_CurrWR:= REAL_TO_WORD(g_stStSysParam.astStUnitParam_UnSave[iN].rHz_UnitScraper_CurrWR *100);
	astStParam_UnitHMI485_Wr_81[iN].wHz_UnitHotWind_CurrWR:= REAL_TO_WORD(g_stStSysParam.astStUnitParam_UnSave[iN].rHz_UnitHotWind_CurrWR*100);
	astStParam_UnitHMI485_Wr_81[iN].wHz_UnitHotWind2_CurrWR:= REAL_TO_WORD(g_stStSysParam.astStUnitParam_UnSave[iN].rHz_UnitHotWind2_CurrWR*100);
	astStParam_UnitHMI485_Wr_81[iN].wPV_UnitTemCtl:= REAL_TO_WORD(g_stStSysParam.astStUnitParam_UnSave[iN].rPV_UnitTemCtl);
	astStParam_UnitHMI485_Wr_81[iN].wSts_UnitTemCtl:= g_stStSysParam.astStUnitParam_UnSave[iN].wSTS_UnitTemCtl;
	astStParam_UnitHMI485_Wr_81[iN].rPos_PrnRoller_Pressure_M:= g_stStSysParam.astStUnitParam_UnSave[iN].rPos_PrnRoller_Pressure_M;
	astStParam_UnitHMI485_Wr_81[iN].rPos_PrnRoller_Pressure_G:= g_stStSysParam.astStUnitParam_UnSave[iN].rPos_PrnRoller_Pressure_G;
	astStParam_UnitHMI485_Wr_81[iN].rPos_NetRoller_Pressure_M:= g_stStSysParam.astStUnitParam_UnSave[iN].rPos_NetRoller_Pressure_M;
	astStParam_UnitHMI485_Wr_81[iN].rPos_NetRoller_Pressure_G:= g_stStSysParam.astStUnitParam_UnSave[iN].rPos_NetRoller_Pressure_G;

	astStParam_UnitHMI485_Wr_82[iN].byPackId:= 2;
	SysMemCmp(ADR(astStParam_UnitHMI485_Wr_82[iN].abyRsv_LowComm),0,SIZEOF(astStParam_UnitHMI485_Wr_82[iN].abyRsv_LowComm));

	IF iN=2 AND astStParam_UnitHMI485_Wr_81[iN].bySts_Ctl.0 THEN(*2色控制1色*)
		iGrpIdTmp:= g_stStSysParam.astStUnitParam_Save[1].byGrpId;
		astStParam_UnitHMI485_Wr_83[iN].byPackId:= 3;
		astStParam_UnitHMI485_Wr_83[iN].wGirth_OtherUnit:= REAL_TO_WORD(g_stStSysParam.astStUnitParam_Save[1].rGirth_Sam*10);
		astStParam_UnitHMI485_Wr_83[iN].iCompanyId_OtherUnit:= g_stStSysParam.stStSysParam_Save.iCustomerId;
		astStParam_UnitHMI485_Wr_83[iN].iPromptMsgId_OtherUnit:= g_stStSysParam.astStGrpParam_UnSave[iGrpIdTmp].iPromptMsg;
		astStParam_UnitHMI485_Wr_83[iN].wAxisId_And_GrpId_OtherUnit:= SHL(INT_TO_WORD(iN),8)+INT_TO_WORD(iGrpIdTmp);
		astStParam_UnitHMI485_Wr_83[iN].wLedtime_And_Language_OtherUnit:= SHL(BYTE_TO_WORD(g_stStSysParam.stStSysParam_Save.byMinutes_ScrSaver),8)+
																	BYTE_TO_WORD(g_stStSysParam.stStSysParam_Save.byLanguageId);
		astStParam_UnitHMI485_Wr_83[iN].iVel_Axis_OtherUnit:= REAL_TO_INT(g_stStSysParam.astStUnitParam_UnSave[1].rAxisVel_PrnRoller*10.0);
		astStParam_UnitHMI485_Wr_83[iN].iVel_Grp_OtherUnit:= REAL_TO_INT(g_stStSysParam.astStGrpParam_UnSave[iGrpIdTmp].rVel_Cur*10.0);
		astStParam_UnitHMI485_Wr_83[iN].wIndex_And_ErrNum_OtherUnit:= g_stStSysParam.astStUnitParam_UnSave[1].byIndex;
		astStParam_UnitHMI485_Wr_83[iN].wUnit_Input_I_OtherUnit:= g_stStSysParam.astStUnitParam_UnSave[1].wUnit_input_I;
		astStParam_UnitHMI485_Wr_83[iN].wUnit_Input_II_OtherUnit:= g_stStSysParam.astStUnitParam_UnSave[1].wUnit_input_II;
		astStParam_UnitHMI485_Wr_83[iN].wUnit_Input_III_OtherUnit:= g_stStSysParam.astStUnitParam_UnSave[1].wUnit_input_III;
		astStParam_UnitHMI485_Wr_83[iN].wHz_UnitInkRoller_CurrWR_OtherUnit:= REAL_TO_WORD(g_stStSysParam.astStUnitParam_UnSave[1].rHz_UnitInkRoller_CurrWR*100);
		astStParam_UnitHMI485_Wr_83[iN].wHz_UnitScraper_CurrWR_OtherUnit:= REAL_TO_WORD(g_stStSysParam.astStUnitParam_UnSave[1].rHz_UnitScraper_CurrWR *100);
		astStParam_UnitHMI485_Wr_83[iN].wHz_UnitHotWind_CurrWR_OtherUnit:= REAL_TO_WORD(g_stStSysParam.astStUnitParam_UnSave[1].rHz_UnitHotWind_CurrWR*100);
		astStParam_UnitHMI485_Wr_83[iN].wHz_UnitHotWind2_CurrWR_OtherUnit:= REAL_TO_WORD(g_stStSysParam.astStUnitParam_UnSave[1].rHz_UnitHotWind2_CurrWR*100);
		astStParam_UnitHMI485_Wr_83[iN].wPV_UnitTemCtl_OtherUnit:= REAL_TO_WORD(g_stStSysParam.astStUnitParam_UnSave[1].rPV_UnitTemCtl);
		astStParam_UnitHMI485_Wr_83[iN].wSts_UnitTemCtl_OtherUnit:= g_stStSysParam.astStUnitParam_UnSave[iN].wSTS_UnitTemCtl;
		astStParam_UnitHMI485_Wr_83[iN].rPos_PrnRoller_Pressure_M_OtherUnit:= g_stStSysParam.astStUnitParam_UnSave[1].rPos_PrnRoller_Pressure_M;
		astStParam_UnitHMI485_Wr_83[iN].rPos_PrnRoller_Pressure_G_OtherUnit:= g_stStSysParam.astStUnitParam_UnSave[1].rPos_PrnRoller_Pressure_G;
		astStParam_UnitHMI485_Wr_83[iN].rPos_NetRoller_Pressure_M_OtherUnit:= g_stStSysParam.astStUnitParam_UnSave[1].rPos_NetRoller_Pressure_M;
		astStParam_UnitHMI485_Wr_83[iN].rPos_NetRoller_Pressure_G_OtherUnit:= g_stStSysParam.astStUnitParam_UnSave[1].rPos_NetRoller_Pressure_G;
	END_IF
(*
	astStParam_UnitHMI485_WrRd[iN].byAxisId:= INT_TO_BYTE(iN);
	astStParam_UnitHMI485_WrRd[iN].iAdjust_V:=
	astStParam_UnitHMI485_WrRd[iN].iAdjust_H:=
	astStParam_UnitHMI485_WrRd[iN].wStatus:= ;
	astStParam_UnitHMI485_WrRd[iN].wUnit_Outout_I:= ;
	astStParam_UnitHMI485_WrRd[iN].wUnit_Outout_II:= ;
*)
END_FOR
